METHOD INTERNAL ParseResponsePayload : DINT
VAR_INPUT
  /// Response data
  ResponseData : RobotLibraryResponseDataFB;
  /// Timestamp
  Timestamp    : SystemTime;  
END_VAR
VAR
  /// Parameter count
 _parameterCnt : DINT;
END_VAR
// Table 6-18: Received CMD payload (RC to PLC) of "ReadRobotData"
// --------------------------
// Header
// --------------------------
// Byte 00 : USINT   - ParSeq | State     
// Byte 01 : SINT    - AlarmMessageSeverity    
// Byte 02 : UINT    - AlarmMessageCode HB
// Byte 03 :         - AlarmMessageCode LB
// --------------------------
// Datablock
// --------------------------
// Byte 04 : CHAR  RCManufacturer[0];
// Byte 05 : CHAR  RCManufacturer[1];
// Byte 06 : CHAR  RCManufacturer[2];
// Byte 07 : CHAR  RCManufacturer[3];
// Byte 08 : CHAR  RCManufacturer[4];
// Byte 09 : CHAR  RCManufacturer[5];
// Byte 10 : CHAR  RCManufacturer[6];
// Byte 11 : CHAR  RCManufacturer[7];
// Byte 12 : CHAR  RCManufacturer[8];
// Byte 13 : CHAR  RCManufacturer[9];
// Byte 14 : CHAR  RCManufacturer[10];
// Byte 15 : CHAR  RCManufacturer[11];
// Byte 16 : CHAR  RCManufacturer[12];
// Byte 17 : CHAR  RCManufacturer[13];
// Byte 18 : CHAR  RCManufacturer[14];
// Byte 19 : CHAR  RCManufacturer[15];
// Byte 20 : CHAR  RCManufacturer[16];
// Byte 21 : CHAR  RCManufacturer[17];
// Byte 22 : CHAR  RCManufacturer[18];
// Byte 23 : CHAR  RCManufacturer[19];
// Byte 24 : CHAR  RCOrderID[0];
// Byte 25 : CHAR  RCOrderID[1];
// Byte 26 : CHAR  RCOrderID[2];
// Byte 27 : CHAR  RCOrderID[3];
// Byte 28 : CHAR  RCOrderID[4];
// Byte 29 : CHAR  RCOrderID[5];
// Byte 30 : CHAR  RCOrderID[6];
// Byte 31 : CHAR  RCOrderID[7];
// Byte 32 : CHAR  RCOrderID[8];
// Byte 33 : CHAR  RCOrderID[9];
// Byte 34 : CHAR  RCOrderID[10];
// Byte 35 : CHAR  RCOrderID[11];
// Byte 36 : CHAR  RCOrderID[12];
// Byte 37 : CHAR  RCOrderID[13];
// Byte 38 : CHAR  RCOrderID[14];
// Byte 39 : CHAR  RCOrderID[15];
// Byte 40 : CHAR  RCOrderID[16];
// Byte 41 : CHAR  RCOrderID[17];
// Byte 42 : CHAR  RCOrderID[18];
// Byte 43 : CHAR  RCOrderID[19];
// Byte 44 : CHAR  RCSerialNumber[0];
// Byte 45 : CHAR  RCSerialNumber[1];
// Byte 46 : CHAR  RCSerialNumber[2];
// Byte 47 : CHAR  RCSerialNumber[3];
// Byte 48 : CHAR  RCSerialNumber[4];
// Byte 49 : CHAR  RCSerialNumber[5];
// Byte 50 : CHAR  RCSerialNumber[6];
// Byte 51 : CHAR  RCSerialNumber[7];
// Byte 52 : CHAR  RCSerialNumber[8];
// Byte 53 : CHAR  RCSerialNumber[9];
// Byte 54 : CHAR  RCSerialNumber[10];
// Byte 55 : CHAR  RCSerialNumber[11];
// Byte 56 : CHAR  RCSerialNumber[12];
// Byte 57 : CHAR  RCSerialNumber[13];
// Byte 58 : CHAR  RCSerialNumber[14];
// Byte 59 : CHAR  RCSerialNumber[15];
// Byte 60 : CHAR  RASerialNumber[0];
// Byte 61 : CHAR  RASerialNumber[1];
// Byte 62 : CHAR  RASerialNumber[2];
// Byte 63 : CHAR  RASerialNumber[3];
// Byte 64 : CHAR  RASerialNumber[4];
// Byte 65 : CHAR  RASerialNumber[5];
// Byte 66 : CHAR  RASerialNumber[6];
// Byte 67 : CHAR  RASerialNumber[7];
// Byte 68 : CHAR  RASerialNumber[8];
// Byte 69 : CHAR  RASerialNumber[9];
// Byte 70 : CHAR  RASerialNumber[10];
// Byte 71 : CHAR  RASerialNumber[11];
// Byte 72 : CHAR  RASerialNumber[12];
// Byte 73 : CHAR  RASerialNumber[13];
// Byte 74 : CHAR  RASerialNumber[14];
// Byte 75 : CHAR  RASerialNumber[15];
// Byte 76 : CHAR  RCFirmwareVersion[0];
// Byte 77 : CHAR  RCFirmwareVersion[1];
// Byte 78 : CHAR  RCFirmwareVersion[2];
// Byte 79 : CHAR  RCFirmwareVersion[3];
// Byte 80 : CHAR  RCFirmwareVersion[4];
// Byte 81 : CHAR  RCFirmwareVersion[5];
// Byte 82 : CHAR  RCFirmwareVersion[6];
// Byte 83 : CHAR  RCFirmwareVersion[7];
// Byte 84 : CHAR  RCFirmwareVersion[8];
// Byte 85 : CHAR  RCFirmwareVersion[9];
// Byte 86 : CHAR  RCFirmwareVersion[10];
// Byte 87 : CHAR  RCFirmwareVersion[11];
// Byte 88 : CHAR  RCInterpreterVersion[0];
// Byte 89 : CHAR  RCInterpreterVersion[1];
// Byte 90 : CHAR  RCInterpreterVersion[2];
// Byte 91 : BYTE  Reserved;
// Byte 92 : BYTE  AxisJointUsed;
// Byte 93 : BYTE  AxisExternalUsed;
// Byte 94 : BYTE  AxisJointUnit;
// Byte 95 : BYTE  AxisExternalUnit;
// Byte 96 : BYTE  RCSupportedFunctions[0];
// Byte 97 : BYTE  RCSupportedFunctions[1];
// Byte 98 : BYTE  RCSupportedFunctions[2];
// Byte 99 : BYTE  RCSupportedFunctions[3];
// Byte 100: BYTE  RCSupportedFunctions[4];
// Byte 101: BYTE  RCSupportedFunctions[5];
// Byte 102: BYTE  RCSupportedFunctions[6];
// Byte 103: BYTE  RCSupportedFunctions[7];
// Byte 104: BYTE  RCSupportedFunctions[8];
// Byte 105: BYTE  RCSupportedFunctions[9];
// Byte 106: BYTE  RCSupportedFunctions[10];
// Byte 107: BYTE  RCSupportedFunctions[11];
// Byte 108: BYTE  RCSupportedFunctions[12];
// Byte 109: BYTE  RCSupportedFunctions[13];
// Byte 110: BYTE  RCSupportedFunctions[14];
// Byte 111: BYTE  RCSupportedFunctions[15];
// Byte 112: BYTE  RCSupportedFunctions[16];
// Byte 113: BYTE  RCSupportedFunctions[17];
// Byte 114: BYTE  RCSupportedFunctions[18];
// Byte 115: BYTE  Reserved;
// Byte 116: CHAR  RobotID[0];
// Byte 117: CHAR  RobotID[1];
// Byte 118: CHAR  RobotID[2];
// Byte 119: CHAR  RobotID[3];
// Byte 120: CHAR  RobotID[4];
// Byte 121: CHAR  RobotID[5];
// Byte 122: CHAR  RobotID[6];
// Byte 123: CHAR  RobotID[7];
// Byte 124: CHAR  RobotID[8];
// Byte 125: CHAR  RobotID[9];
// Byte 126: CHAR  RobotID[10];
// Byte 127: CHAR  RobotID[11];
// Byte 128: CHAR  RobotID[12];
// Byte 129: CHAR  RobotID[13];
// Byte 130: CHAR  RobotID[14];
// Byte 131: CHAR  RobotID[15];
// Byte 132: UINT  InterpreterCycleTime HW HB;
// Byte 133:       InterpreterCycleTime HW LB;
// --------------------------

                  
                  // call base implementation to parse the header from payload buffer
ResponseData.PayloadPtr := SUPER^.ParseResponsePayload(ResponseData := ResponseData, Timestamp := Timestamp);

// ST-FIX F100: missing (trailing zero) bytes of the payload are 0, no values of the previous response
SysDepMemSet( pDest := ADR(_response), Value := 0, DataLen := SIZEOF(_response));

// copy parsed header to response
_response.ParSeq               := _rspHeader.ParSeq;
_response.State                := _rspHeader.State;
_response.AlarmMessageSeverity := _rspHeader.AlarmMessageSeverity;
_response.AlarmMessageCode     := _rspHeader.AlarmMessageCode;


// Check payload remaining ? 
IF ( ResponseData.IsPayloadRemaining)
THEN  
  // Get _response.RCManufacturer
  ResponseData.GetDataBlock(pData := ADR(_response.RCManufacturer)      , SIZEOF(_response.RCManufacturer   )   , IsString := TRUE );
  // inc parameter counter
 _parameterCnt := _parameterCnt + 1;
END_IF


// Check payload remaining ? 
IF ( ResponseData.IsPayloadRemaining)
THEN  
  // Get _response.RCOrderID
  ResponseData.GetDataBlock(pData := ADR(_response.RCOrderID)           , SIZEOF(_response.RCOrderID        )   , IsString := TRUE );
  // inc parameter counter
 _parameterCnt := _parameterCnt + 1;
END_IF


// Check payload remaining ? 
IF ( ResponseData.IsPayloadRemaining)
THEN  
  // Get _response.RCSerialNumber
  ResponseData.GetDataBlock(pData := ADR(_response.RCSerialNumber)      , SIZEOF(_response.RCSerialNumber   )   , IsString := TRUE );
  // inc parameter counter
 _parameterCnt := _parameterCnt + 1;
END_IF


// Check payload remaining ? 
IF ( ResponseData.IsPayloadRemaining)
THEN  
  // Get _response.RASerialNumber
  ResponseData.GetDataBlock(pData := ADR(_response.RASerialNumber)      , SIZEOF(_response.RASerialNumber   )   , IsString := TRUE );
  // inc parameter counter
 _parameterCnt := _parameterCnt + 1;
END_IF


// Check payload remaining ? 
IF ( ResponseData.IsPayloadRemaining)
THEN  
  // Get _response.RCFirmwareVersion
  ResponseData.GetDataBlock(pData := ADR(_response.RCFirmwareVersion)   , SIZEOF(_response.RCFirmwareVersion)   , IsString := TRUE );
  // inc parameter counter
 _parameterCnt := _parameterCnt + 1;
END_IF


// Check payload remaining ? 
IF ( ResponseData.IsPayloadRemaining)
THEN  
  // Get _response.RCInterpreterVersion
  // ResponseData.GetDataBlock(pData := ADR(_response.RCInterpreterVersion), SIZEOF(_response.RCInterpreterVersion), IsString := TRUE );

  // This adaption was made because of Stäubli - check with other robot brands...
  
  // Get _response.RCInterpreterVersion
 // ST-FIX F163: the three numbers, the text is made of them
   _response.RCInterpreterVersionNumber.MajorVersion := BYTE_TO_USINT(ResponseData.GetByte());
   _response.RCInterpreterVersionNumber.MinorVersion := BYTE_TO_USINT(ResponseData.GetByte());
   _response.RCInterpreterVersionNumber.PatchVersion := BYTE_TO_USINT(ResponseData.GetByte());
   _response.RCInterpreterVersion := CONCAT(USINT_TO_STRING(_response.RCInterpreterVersionNumber.MajorVersion), '.');
   _response.RCInterpreterVersion := CONCAT(_response.RCInterpreterVersion, USINT_TO_STRING(_response.RCInterpreterVersionNumber.MinorVersion));
   _response.RCInterpreterVersion := CONCAT(_response.RCInterpreterVersion, '.');
   _response.RCInterpreterVersion := CONCAT(_response.RCInterpreterVersion, USINT_TO_STRING(_response.RCInterpreterVersionNumber.PatchVersion));

  // inc parameter counter
 _parameterCnt := _parameterCnt + 1;
END_IF


// Check payload remaining ? 
IF ( ResponseData.IsPayloadRemaining)
THEN  
  // Get _response.Reserve
 _response.Reserve := ResponseData.GetByte(); 
  // inc parameter counter
 _parameterCnt := _parameterCnt + 1;
END_IF


// Check payload remaining ? 
IF ( ResponseData.IsPayloadRemaining)
THEN  
  // Get _response.AxisJointUsed
 _response.AxisJointUsed := ResponseData.GetByte(); 
  // inc parameter counter
 _parameterCnt := _parameterCnt + 1;
END_IF


// Check payload remaining ? 
IF ( ResponseData.IsPayloadRemaining)
THEN  
  // Get _response.AxisExternalUsed
 _response.AxisExternalUsed := ResponseData.GetByte(); 
  // inc parameter counter
 _parameterCnt := _parameterCnt + 1;
END_IF


// Check payload remaining ? 
IF ( ResponseData.IsPayloadRemaining)
THEN  
  // Get _response.AxisJointUnit
 _response.AxisJointUnit := ResponseData.GetByte(); 
  // inc parameter counter
 _parameterCnt := _parameterCnt + 1;
END_IF


// Check payload remaining ? 
IF ( ResponseData.IsPayloadRemaining)
THEN  
  // Get _response.AxisExternalUnit
 _response.AxisExternalUnit := ResponseData.GetByte();
  // inc parameter counter
 _parameterCnt := _parameterCnt + 1;
END_IF


// Check payload remaining ? 
IF ( ResponseData.IsPayloadRemaining)
THEN  
  // Get _response.RCSupportedFunctions
  ResponseData.GetDataBlock(pData := ADR(_response.RCSupportedFunctions), SIZEOF(_response.RCSupportedFunctions), IsString := FALSE );
  // inc parameter counter
 _parameterCnt := _parameterCnt + 1;
END_IF


// Check payload remaining ? 
IF ( ResponseData.IsPayloadRemaining)
THEN  
  // Get _response.Reserve2
 _response.Reserve2 := ResponseData.GetByte(); 
  // inc parameter counter
 _parameterCnt := _parameterCnt + 1;
END_IF


// Check payload remaining ? 
IF ( ResponseData.IsPayloadRemaining)
THEN  
  // Get _response.RobotID
  ResponseData.GetDataBlock(pData := ADR(_response.RobotID)             , SIZEOF(_response.RobotID)             , IsString := TRUE );
  // inc parameter counter
 _parameterCnt := _parameterCnt + 1;
END_IF


// Check payload remaining ? 
IF ( ResponseData.IsPayloadRemaining)
THEN  
  // Get _response.InterpreterCycleTime
 _response.InterpreterCycleTime := ResponseData.GetUint(); // ST-FIX F30 
  // inc parameter counter
 _parameterCnt := _parameterCnt + 1;
END_IF

 
// Create logging
ParseResponsePayloadLog(ResponseData := ResponseData, Timestamp := Timestamp, ParameterCnt := _parameterCnt);
END_METHOD

METHOD INTERNAL ParseResponsePayloadLog
VAR_INPUT
  /// Response data
  ResponseData : RobotLibraryResponseDataFB;
  /// Timestamp
  Timestamp    : SystemTime;  
  /// Parameter count
  ParameterCnt : DINT;
END_VAR
VAR 
  /// internal index for loops
 _idx : DINT;
  /// temporary string
 _tmpStr : STRING;
END_VAR
// Create log entry for Parameter start
CreateLogMessagePara1 ( Timestamp   := Timestamp,
                        MessageType := MessageType.CMD,
                        Severity    := Severity.DEBUG,
                        MessageCode := 0,
                        MessageText := '{1} parameter(s) to parse from the response data:',
                        Para1       := DINT_TO_STRING(ParameterCnt));


// Return if no parameter is remaining...
IF ( ParameterCnt = 0 ) THEN RETURN; END_IF
// dec remaining parameter(s)                        
ParameterCnt := ParameterCnt - 1;
// Create log entry for RCManufacturer
CreateLogMessagePara1 ( Timestamp   := Timestamp,
                        MessageType := MessageType.CMD,
                        Severity    := Severity.DEBUG,
                        MessageCode := 0,
                        MessageText := 'Response.RCManufacturer = {1}',
                        Para1       := _response.RCManufacturer);


// Return if no parameter is remaining...
IF ( ParameterCnt = 0 ) THEN RETURN; END_IF
// dec remaining parameter(s)                        
ParameterCnt := ParameterCnt - 1;
// Create log entry for RCOrderID
CreateLogMessagePara1 ( Timestamp   := Timestamp,
                        MessageType := MessageType.CMD,
                        Severity    := Severity.DEBUG,
                        MessageCode := 0,
                        MessageText := 'Response.RCOrderID = {1}',
                        Para1       := _response.RCOrderID);


// Return if no parameter is remaining...
IF ( ParameterCnt = 0 ) THEN RETURN; END_IF
// dec remaining parameter(s)                        
ParameterCnt := ParameterCnt - 1;
// Create log entry for RCSerialNumber
CreateLogMessagePara1 ( Timestamp   := Timestamp,
                        MessageType := MessageType.CMD,
                        Severity    := Severity.DEBUG,
                        MessageCode := 0,
                        MessageText := 'Response.RCSerialNumber = {1}',
                        Para1       := _response.RCSerialNumber);


// Return if no parameter is remaining...
IF ( ParameterCnt = 0 ) THEN RETURN; END_IF
// dec remaining parameter(s)                        
ParameterCnt := ParameterCnt - 1;
// Create log entry for RASerialNumber
CreateLogMessagePara1 ( Timestamp   := Timestamp,
                        MessageType := MessageType.CMD,
                        Severity    := Severity.DEBUG,
                        MessageCode := 0,
                        MessageText := 'Response.RASerialNumber = {1}',
                        Para1       := _response.RASerialNumber);


// Return if no parameter is remaining...
IF ( ParameterCnt = 0 ) THEN RETURN; END_IF
// dec remaining parameter(s)                        
ParameterCnt := ParameterCnt - 1;
// Create log entry for RCFirmwareVersion
CreateLogMessagePara1 ( Timestamp   := Timestamp,
                        MessageType := MessageType.CMD,
                        Severity    := Severity.DEBUG,
                        MessageCode := 0,
                        MessageText := 'Response.RCFirmwareVersion = {1}',
                        Para1       := _response.RCFirmwareVersion);
                        

// Return if no parameter is remaining...
IF ( ParameterCnt = 0 ) THEN RETURN; END_IF
// dec remaining parameter(s)                        
ParameterCnt := ParameterCnt - 1;
// Create log entry for RCInterpreterVersion
CreateLogMessagePara1 ( Timestamp   := Timestamp,
                        MessageType := MessageType.CMD,
                        Severity    := Severity.DEBUG,
                        MessageCode := 0,
                        MessageText := 'Response.RCInterpreterVersion = {1}',
                        Para1       := _response.RCInterpreterVersion);


// Return if no parameter is remaining...
IF ( ParameterCnt = 0 ) THEN RETURN; END_IF
// dec remaining parameter(s)                        
ParameterCnt := ParameterCnt - 1;
// Create log entry for Reserve
CreateLogMessagePara1 ( Timestamp   := Timestamp,
                        MessageType := MessageType.CMD,
                        Severity    := Severity.DEBUG,
                        MessageCode := 0,
                        MessageText := 'Response.Reserve = {1}',
                        Para1       :=  BYTE_TO_STRING(_response.Reserve));


// Return if no parameter is remaining...
IF ( ParameterCnt = 0 ) THEN RETURN; END_IF
// dec remaining parameter(s)                        
ParameterCnt := ParameterCnt - 1;
// Create log entry for AxisJointUsed
CreateLogMessagePara1 ( Timestamp   := Timestamp,
                        MessageType := MessageType.CMD,
                        Severity    := Severity.DEBUG,
                        MessageCode := 0,
                        MessageText := 'Response.AxisJointUsed = {1}',
                        Para1       :=  BYTE_TO_STRING_BIN(_response.AxisJointUsed));


// Return if no parameter is remaining...
IF ( ParameterCnt = 0 ) THEN RETURN; END_IF
// dec remaining parameter(s)                        
ParameterCnt := ParameterCnt - 1;
// Create log entry for AxisExternalUsed
CreateLogMessagePara1 ( Timestamp   := Timestamp,
                        MessageType := MessageType.CMD,
                        Severity    := Severity.DEBUG,
                        MessageCode := 0,
                        MessageText := 'Response.AxisExternalUsed = {1}',
                        Para1       :=  BYTE_TO_STRING_BIN(_response.AxisExternalUsed));


// Return if no parameter is remaining...
IF ( ParameterCnt = 0 ) THEN RETURN; END_IF
// dec remaining parameter(s)                        
ParameterCnt := ParameterCnt - 1;
// Create log entry for AxisJointUnit
CreateLogMessagePara1 ( Timestamp   := Timestamp,
                        MessageType := MessageType.CMD,
                        Severity    := Severity.DEBUG,
                        MessageCode := 0,
                        MessageText := 'Response.AxisJointUnit = {1}',
                        Para1       :=  BYTE_TO_STRING(_response.AxisJointUnit));


// Return if no parameter is remaining...
IF ( ParameterCnt = 0 ) THEN RETURN; END_IF
// dec remaining parameter(s)                        
ParameterCnt := ParameterCnt - 1;
// Create log entry for AxisExternalUnit
CreateLogMessagePara1 ( Timestamp   := Timestamp,
                        MessageType := MessageType.CMD,
                        Severity    := Severity.DEBUG,
                        MessageCode := 0,
                        MessageText := 'Response.AxisExternalUnit = {1}',
                        Para1       :=  BYTE_TO_STRING(_response.AxisExternalUnit));

FOR _idx := 0 TO 18
do
 _tmpStr := '2#';
 _tmpStr := CONCAT( _tmpStr, BYTE_TO_STRING_BIN(_response.RCSupportedFunctions[_idx]));

  // Return if no parameter is remaining...
  IF ( ParameterCnt = 0 ) THEN RETURN; END_IF
  // dec remaining parameter(s)                        
  ParameterCnt := ParameterCnt - 1;
  // Create log entry for RCSupportedFunctions
  CreateLogMessagePara2 ( Timestamp   := Timestamp,
                          MessageType := MessageType.CMD,
                          Severity    := Severity.DEBUG,
                          MessageCode := 0,
                          MessageText := 'Response.RCSupportedFunctions[{2}] = {1}',
                          Para1       := _tmpStr,
                          Para2       :=  DINT_TO_STRING(_idx));
END_FOR


// Return if no parameter is remaining...
IF ( ParameterCnt = 0 ) THEN RETURN; END_IF
// dec remaining parameter(s)                        
ParameterCnt := ParameterCnt - 1;
// Create log entry for Reserve2
CreateLogMessagePara1 ( Timestamp   := Timestamp,
                        MessageType := MessageType.CMD,
                        Severity    := Severity.DEBUG,
                        MessageCode := 0,
                        MessageText := 'Response.Reserve2 = {1}',
                        Para1       :=  BYTE_TO_STRING(_response.Reserve2));


// Return if no parameter is remaining...
IF ( ParameterCnt = 0 ) THEN RETURN; END_IF
// dec remaining parameter(s)                        
ParameterCnt := ParameterCnt - 1;
// Create log entry for RobotID
CreateLogMessagePara1 ( Timestamp   := Timestamp,
                        MessageType := MessageType.CMD,
                        Severity    := Severity.DEBUG,
                        MessageCode := 0,
                        MessageText := 'Response.RobotID = {1}',
                        Para1       :=  _response.RobotID);


// Return if no parameter is remaining...
IF ( ParameterCnt = 0 ) THEN RETURN; END_IF
// dec remaining parameter(s)                        
ParameterCnt := ParameterCnt - 1;
// Create log entry for InterpreterCycleTime
CreateLogMessagePara1 ( Timestamp   := Timestamp,
                        MessageType := MessageType.CMD,
                        Severity    := Severity.DEBUG,
                        MessageCode := 0,
                        MessageText := 'Response.InterpreterCycleTime = {1}',
                        Para1       :=  UINT_TO_STRING(_response.InterpreterCycleTime));
END_METHOD

METHOD PROTECTED Reset : DINT
VAR_INPUT
END_VAR
Reset := SUPER^.Reset();

Done               := FALSE;
Busy               := FALSE;
CommandBuffered    := FALSE;
END_METHOD

END_FUNCTION_BLOCK

// Library/POUs/_internal/BaseFBs/RobotLibraryBaseExecuteFB
FUNCTION_BLOCK RobotLibraryBaseExecuteFB EXTENDS RobotLibraryBaseFB
// ------------------------------------------------------------------------- 
//  SRCI Robot Library                                                
// ------------------------------------------------------------------------- 
//                                                                           
//  Object:      RobotLibraryBaseFB                                       
//  Author:      Thorsten Brach                                                
//  Date:        2024-08-11
//
//  Description:                                              
//   
//                                                                           
//  Copyright: 
//    (C) 2024 Thorsten Brach. All rights reserved                                                                                                                                            
//             Licensed under the MIT License.
//                                                                           
//  Disclaimer:                                                                           
//    This project is provided without any guarantee and can be used for   
//    private and commercial purposes. Any use is at the user’s 
//    own risk and responsibility.
//
// -------------------------------------------------------------------------
VAR_INPUT
  /// Start of the command at the rising edge
  Execute         : BOOL;
END_VAR
VAR_OUTPUT
  /// The command has been completed successfully
  Done            : BOOL;
  /// FB is being processed
  Busy            : BOOL;
  /// Command is transferred and confirmed by the RC
//  CommandBuffered : BOOL;  
END_VAR


VAR
  /// Rising edge for execute
  {attribute 'hide'}
 _execute_R       : R_TRIG;
  /// Falling edge for execute
  {attribute 'hide'}
 _execute_F       : F_TRIG;
END_VAR
            
          
VAR
  _executeIn : BOOL;
  _executeHold : BOOL;
END_VAR
VAR
  /// ST-FIX F104: rising edge of the Execute input (also while Busy)
  _executeRestart_R : R_TRIG;
END_VAR

// ST-FIX F50: a falling edge of Execute must not cancel the command (spec 5.5.x "Output
// status"): Execute is held internally while Busy; Done/Error/CommandAborted of a command
// whose Execute is already FALSE are shown for one cycle, then the block resets
_executeIn := Execute;
// ST-FIX F104: rising edge of the Execute input also while Busy (Execute is held, F50)
_executeRestart_R(CLK := Execute);
Execute     := Execute OR _executeHold;
SUPER^(AxesGroup := AxesGroup);
_executeHold := Busy;
Execute      := _executeIn;

// Base implementation must be called ! 
METHOD PROTECTED OnCall
VAR_IN_OUT
  /// Robot assignment of function
  AxesGroup         : AxesGroup; 
END_VAR

VAR
  /// internal return value
 _retVal : DINT;
END_VAR
SUPER^.OnCall(AxesGroup := AxesGroup);

// building rising and falling edges
_execute_R( CLK := Execute);
_execute_F( CLK := Execute);


// Check command execution is allowed ?
IF ((     Execute                                ) AND
    ( NOT AxesGroup.State.CMDsEnabled            ) AND
    (     MyType <> 'MC_ExchangeConfigurationFB' ) AND // is part of init sequence
    (     MyType <> 'MC_ReadMessagesFB'          ) AND // is part of init sequence
    (     MyType <> 'MC_ReadRobotDataFB'         ))    // is part of init sequence
THEN
  SetError( ErrorID := RobotLibraryErrorIdEnum.ERR_COMMANDS_NOT_ENABLED, Overwrite := TRUE );
  Error   := TRUE;
  Busy    := FALSE;
END_IF


// On execution started
IF ( _execute_R.Q )
THEN
  OnExecStart(AxesGroup := AxesGroup);
END_IF


// On execution cancel  
IF ( Busy ) AND ( _execute_F.Q ) 
THEN
  // set cancel flag
 _cancel := TRUE;
END_IF

IF ( _cancel )
THEN
  // call Cancel
 _retVal := OnExecCancel(AxesGroup := AxesGroup);
  
  // done or error ?
  IF ( _retVal <> RobotLibraryConstants.RUNNING )
  THEN
    // reset cancel flag
   _cancel := FALSE;
	END_IF
END_IF


// On execution error clear
IF ( Error ) AND ( _execute_F.Q )
THEN
  // set ClearError flag
 _clearError := TRUE;
END_IF

IF ( _clearError )
THEN
 _retVal := OnExecErrorClear(AxesGroup := AxesGroup); 

  // done or error ?
  IF ( _retVal <> RobotLibraryConstants.RUNNING )
  THEN
    // reset ClearError flag
   _clearError := FALSE;
	END_IF
END_IF
END_METHOD

METHOD PROTECTED OnExecCancel : DINT
VAR_IN_OUT
  /// Robot assignment of function
  AxesGroup : AxesGroup; 
END_VAR
VAR
  /// internal return value 
 _retVal    : DINT;
END_VAR
// Create log entry
CreateLogMessagePara1 ( Timestamp   := AxesGroup.State.SystemTime,
                        MessageType := MessageType.CMD,
                        Severity    := Severity.DEBUG,
                        MessageCode := 0,
                        MessageText := 'Execution of {1} cancled ',
                        Para1       := MyType);                 

// try to remove cmd
_retVal := AxesGroup.Acyclic.ActiveCommandRegister.RemoveCmd(_uniqueID);


IF (_retVal = RobotLibraryConstants.OK)
THEN
  // Create log entry
  CreateLogMessagePara1 ( Timestamp   := AxesGroup.State.SystemTime,
                          MessageType := MessageType.CMD,
                          Severity    := Severity.DEBUG,
                          MessageCode := 0,
                          MessageText := '{1} successfully removed from ACR',
                          Para1       := MyType);                 
ELSE
  // Create log entry
  CreateLogMessagePara1 ( Timestamp   := AxesGroup.State.SystemTime,
                          MessageType := MessageType.CMD,
                          Severity    := Severity.DEBUG,
                          MessageCode := 0,
                          MessageText := '{1} was not removed from ACR because execution was already in progress',
                          Para1       := MyType);                 
END_IF


OnExecCancel := Reset();
END_METHOD

METHOD PROTECTED OnExecErrorClear : DINT
VAR_IN_OUT
  /// Robot assignment of function
  AxesGroup : AxesGroup; 
END_VAR
OnExecErrorClear := Reset();
END_METHOD

METHOD PROTECTED OnExecRun : DINT
VAR_IN_OUT
  /// Robot assignment of function
  AxesGroup : AxesGroup; 
END_VAR
END_METHOD

METHOD PROTECTED OnExecStart : DINT
VAR_IN_OUT
  /// Robot assignment of function
  AxesGroup : AxesGroup; 
END_VAR


// ST-FIX F71: Priority (1 = very high ... 4 = low, table 7-1)
IF ( Priority < PriorityLevel.VERY_HIGH )
THEN
  SetError( ErrorID := RobotLibraryErrorIdEnum.ERR_PRIORITY_TOO_HIGH, Overwrite := TRUE );
  // Create log entry
  CreateLogMessage ( Timestamp   := AxesGroup.State.SystemTime,
                     MessageType := MessageType.CMD,
                     Severity    := Severity.ERROR,
                     MessageCode := ErrorID,
                     MessageText := 'Invalid input Priority: higher than VERY_HIGH');
  Error := TRUE;
ELSIF ( Priority > PriorityLevel.LOW )
THEN
  SetError( ErrorID := RobotLibraryErrorIdEnum.ERR_PRIORITY_TOO_LOW, Overwrite := TRUE );
  // Create log entry
  CreateLogMessage ( Timestamp   := AxesGroup.State.SystemTime,
                     MessageType := MessageType.CMD,
                     Severity    := Severity.ERROR,
                     MessageCode := ErrorID,
                     MessageText := 'Invalid input Priority: lower than LOW');
  Error := TRUE;
END_IF
END_METHOD

METHOD PROTECTED OnUpdateStateFlags
VAR_INPUT
  /// Command message state
  State : CmdMessageState;
END_VAR
// Reset State flags
Done := FALSE;

CASE State OF

  // No operation or process is active
  CmdMessageState.EMPTY               :;
  // Created but not yet started
  CmdMessageState.CREATED             :;
  // Buffered and awaiting execution
  CmdMessageState.BUFFERED            :;
  // Buffered in planner for future execution
  CmdMessageState.BUFFERED_IN_PLANNER :;
  // Currently active and in progress
  CmdMessageState.ACTIVE              :;
  // Interrupted and awaiting continuation
  CmdMessageState.INTERRUPTED         :;
  // Requested for abort
  CmdMessageState.ABORT_REQUEST       :;
  // Successfully completed
  CmdMessageState.DONE                : Done := TRUE;
                                        Busy := FALSE;
  // Aborted before completion
  CmdMessageState.ABORTED             : Busy := FALSE;
  // Encountered an error during execution
  CmdMessageState.ERROR               : Error := TRUE;
                                        Busy  := FALSE;
END_CASE
END_METHOD

METHOD PROTECTED Reset : DINT
VAR_INPUT
END_VAR
Reset := SUPER^.Reset();

Done := FALSE;
Busy := FALSE;
END_METHOD

END_FUNCTION_BLOCK

// Library/POUs/_internal/LogFBs/AxesGroupMessageLogFB
FUNCTION_BLOCK AxesGroupMessageLogFB IMPLEMENTS IMessageLogger
// ------------------------------------------------------------------------- 
//  SRCI Robot Library                                                
// ------------------------------------------------------------------------- 
//                                                                           
//  Object:      AxesGroupMessageLogFB                                       
//  Author:      Thorsten Brach                                                
//  Date:        2025-01-05
//
//  Description:                                              
//   
//                                                                           
//  Copyright: 
//    (C) 2025 Thorsten Brach. All rights reserved                                                                                                                                            
//             Licensed under the MIT License.
//                                                                           
//  Disclaimer:                                                                           
//    This project is provided without any guarantee and can be used for   
//    private and commercial purposes. Any use is at the user’s 
//    own risk and responsibility.
//
// -------------------------------------------------------------------------
VAR_INPUT
  /// Logging level
  LogLevel         : LogLevel;
  /// Interface to an external logger
  ExternalLogger   : IMessageLogger;
END_VAR


VAR_OUTPUT
  /// Amount of system log entries
  SystemLogEntries : UINT := 0;
  /// Amount of message log entries
  MessagesEntries  : UINT := 0;
  /// System log
  SystemLogs       : ARRAY[0..RobotLibraryParameter.SYSTEM_LOG_MAX ] OF STRING(RobotLibraryParameter.MESSAGE_TEXT_LEN);
  /// Message Log
  Messages         : ARRAY[0..RobotLibraryParameter.MESSAGE_LOG_MAX] OF AlarmMessage;  
END_VAR

METHOD PUBLIC AddMessageLog
VAR_INPUT
  MessageLog : AlarmMessage;
END_VAR

VAR
  /// internal index
 _idx            : DINT;
  /// internal index to delete
 _idxFound       : DINT;
  /// lowest Severity
 _lowestSeverity : Severity := Severity.FATAL_ERROR;
  /// temporary buffer ( must be one element less than the message log !!! )
 _tmpBuffer      : ARRAY[0..RobotLibraryParameter.MESSAGE_LOG_MAX -1] OF AlarmMessage; 
END_VAR

                  // Check entry must be added ? 
IF (( LogLevel  <= MessageLog.Severity     ) AND
    ( LogLevel  >  LogLevelEnum.DEACTIVATE ))
THEN
  // Check message buffer is full ? 
  IF ( MessagesEntries >= RobotLibraryParameter.MESSAGE_LOG_MAX )
  THEN
    // find lowest Severity
    FOR _idx := 1 TO RobotLibraryParameter.MESSAGE_LOG_MAX
    DO
      // check entry has a lower severity ? 
     _lowestSeverity := MIN( Messages[_idx].Severity, _lowestSeverity );
		END_FOR

    // search for the oldes message with a lower Severity 
    FOR _idx := RobotLibraryParameter.MESSAGE_LOG_MAX TO 1 BY -1
    DO
      // message found ?
      IF (( Messages[_idx].Severity <   MessageLog.Severity ) AND
          ( Messages[_idx].Severity <= _lowestSeverity      ))
      THEN
        // save index to delete 
       _idxFound := _idx;
        EXIT;
			END_IF
		END_FOR
    
    // check message must be deleted ? 
    IF ( _idxFound > 0 )
    THEN
      // shift all messages starting from the found index one position forwards
      FOR _idx := _idxFound TO RobotLibraryParameter.MESSAGE_LOG_MAX -1
      DO
        Messages[_idx] := Messages[_idx +1];
			END_FOR
		END_IF
  END_IF  

  // shift all messages one position backwards
  // shift messages log entries
  SysDepMemCpy( pDest := ADR(_tmpBuffer[0]), pSrc := ADR(  Messages[0]), DataLen := SIZEOF(_tmpBuffer));
  SysDepMemCpy( pDest := ADR(  Messages[1]), pSrc := ADR(_tmpBuffer[0]), DataLen := SIZEOF(_tmpBuffer));
  
  
  // Add new message 
  Messages[0].Timestamp   := MessageLog.Timestamp;           
  Messages[0].MessageType := MessageLog.MessageType;
  Messages[0].Severity    := MessageLog.Severity;
  Messages[0].MessageText := MessageLog.MessageText;
  Messages[0].MessageCode := MessageLog.MessageCode;
  Messages[0].AcrID       := MessageLog.AcrID;   // ST-FIX F74
  Messages[0].CmdType     := MessageLog.CmdType; // ST-FIX F74
  
  // inc message counter
  MessagesEntries := DINT_TO_UINT(LIMIT(0, MessagesEntries + 1, RobotLibraryParameter.MESSAGE_LOG_MAX));
END_IF
END_METHOD

METHOD Public AddMessageLogByParameter
VAR_INPUT
  /// Timestamp
  Timestamp   : SystemTime;
  /// Type of message according to Table 5-48:
  MessageType : MessageType;
  /// Severity of message according to Table 5-49: Debug, Info, Warning, Error, Fatal error
  Severity    : Severity;
  /// Code of messages
  MessageCode : DWORD;
  /// Static text of message
  MessageText : STRING(RobotLibraryParameter.MESSAGE_TEXT_LEN);    
END_VAR

VAR
  /// temporary message 
 _message : AlarmMessage;
END_VAR
_message.Timestamp   := Timestamp;
_message.MessageType := MessageType;
_message.MessageCode := MessageCode;
_message.MessageText := MessageText;
_message.Severity    := Severity;

// Add message to message buffer       
AddMessageLog(_message);
END_METHOD

METHOD PUBLIC AddSystemLog
VAR_INPUT
  /// system log message
  SystemLog : STRING(255);
END_VAR
VAR
  /// internal index
 _idx       : DINT;
  /// internal log message 
 _message   : AlarmMessage;
  /// temporary buffer ( must be one element less than the system log !!! )
 _tmpBuffer : ARRAY[0..RobotLibraryParameter.SYSTEM_LOG_MAX -1] OF STRING(RobotLibraryParameter.MESSAGE_TEXT_LEN);
END_VAR
// shift system log entries
SysDepMemCpy( pDest := ADR(_tmpBuffer[0]), pSrc := ADR(SystemLogs[0]), DataLen := SIZEOF(_tmpBuffer));
SysDepMemCpy( pDest := ADR(SystemLogs[1]), pSrc := ADR(_tmpBuffer[0]), DataLen := SIZEOF(_tmpBuffer));

// Delete CR from system log message
SystemLog := StrReplace(SystemLog, '$R', '');
// Delete LF from system log message          
SystemLog := StrReplace(SystemLog, '$N', '');    
       
// Add System log to buffer 
SystemLogs[0] := SystemLog;
 
// inc SystemLog counter
SystemLogEntries := DINT_TO_UINT(LIMIT(0, SystemLogEntries + 1, RobotLibraryParameter.SYSTEM_LOG_MAX));
END_METHOD

METHOD CheckMessageCodePresent : BOOL
VAR_INPUT
  /// Code of messages
  MessageCode : DWORD;
END_VAR

VAR
  /// internal index for loops
 _idx : DINT;
END_VAR
FOR _idx := 0 TO RobotLibraryParameter.MESSAGE_LOG_MAX
DO
  IF (Messages[_idx].MessageCode = MessageCode)
  THEN
    CheckMessageCodePresent := TRUE;
    RETURN;
	END_IF
END_FOR
END_METHOD

METHOD PUBLIC DeleteMessages
VAR_INPUT
END_VAR
// reset messages
SysDepMemSet(ADR(Messages), 0, SIZEOF(Messages));
// reset message counter
MessagesEntries := 0;
END_METHOD

METHOD DeleteSystemLogs
VAR_INPUT
END_VAR
// reset SystemLogs
SysDepMemSet(ADR(SystemLogs), 0, SIZEOF(SystemLogs));
// reset SystemLogs counter
SystemLogEntries := 0;
END_METHOD

END_FUNCTION_BLOCK

// Library/POUs/_internal/SystemData/AxesGroupSystemDataFB
FUNCTION_BLOCK AxesGroupSystemDataFB 
{attribute 'pack_mode' := '1'} 
// ------------------------------------------------------------------------- 
//  SRCI Robot Library                                                
// ------------------------------------------------------------------------- 
//                                                                           
//  Object:      AxesGroupSystemDataFB                                       
//  Author:      Thorsten Brach                                                
//  Date:        2025-08-31
//
//  Description:                                              
//   
//                                                                           
//  Copyright: 
//    (C) 2025 Thorsten Brach. All rights reserved                                                                                                                                            
//             Licensed under the MIT License.
//                                                                           
//  Disclaimer:                                                                           
//    This project is provided without any guarantee and can be used for   
//    private and commercial purposes. Any use is at the user’s 
//    own risk and responsibility.
//
// -------------------------------------------------------------------------
VAR_INPUT
  /// Pointer to ToolData array
  ToolDataPtr       : POINTER TO Tool;
  /// Lower dimension of ToolData array 
  ToolDataMin       : DINT;
  /// Lower dimension of ToolData array
  ToolDataMax       : DINT;
  /// Amount of ToolData elements in array
  ToolDataCount     : UDINT;

  /// Pointer to LoadData array
  LoadDataPtr       : POINTER TO Load;
  /// Lower dimension of LoadData array 
  LoadDataMin       : DINT;
  /// Lower dimension of LoadData array
  LoadDataMax       : DINT;
  /// Amount of Load elements in array
  LoadDataCount     : UDINT;

  /// Pointer to FrameData array
  FrameDataPtr      : POINTER TO Frame;
  /// Lower dimension of FrameData array 
  FrameDataMin      : DINT;
  /// Lower dimension of FrameData array
  FrameDataMax      : DINT;
  /// Amount of FrameData elements in array
  FrameDataCount    : UDINT;
  
  /// Pointer to WorkAreas array
  WorkAreasPtr      : POINTER TO RobotWorkArea;
  /// Lower dimension of WorkAreas array 
  WorkAreasMin      : DINT;
  /// Lower dimension of WorkAreas array
  WorkAreasMax      : DINT;
  /// Amount of WorkAreas elements in array
  WorkAreasCount    : UDINT;
  
  /// Software limits stored on PLC
  SWLimits          : REFERENCE TO SWLimits;
  /// Default dynamics stored on PLC. For more information refer to 5.5.7
  DefaultDynamics   : REFERENCE TO DefaultDynamics;
  /// Reference dynamics stored on PLC. For more information refer to 5.5.7
  ReferenceDynamics : REFERENCE TO ReferenceDynamics;
END_VAR

METHOD UpdateDefaultDynamics : DINT
VAR_INPUT
  /// Default dynamics values according to Table 6-172.
  DynamicValues : DefaultDynamics;
END_VAR
// Check pointer is vaild ?
IF ( NOT __ISVALIDREF(DefaultDynamics))  
THEN
  RETURN;
END_IF

// Applay new values
DefaultDynamics := DynamicValues;
END_METHOD

METHOD UpdateFrameData : DINT
VAR_INPUT
  /// Reference to BaseFB 
  Caller     : REFERENCE TO RobotLibraryBaseFB;
  /// Current System Time
  SystemTime : SystemTime;
  /// Frame index M
  /// • 0: WCS (default) O
  /// • 1..254: UCS (User frames)
  FrameNo    : USINT;
  /// Frame data (see chapter 5.5.6.2)
  FrameData  : FrameData;
END_VAR


VAR
  /// pointer to frame data
  pFrameData : POINTER TO Frame;  
END_VAR
// Check pointer is vaild ?
IF ( FrameDataPtr = RobotLibraryConstants.NULL_POINTER )
THEN
  RETURN;
END_IF

// Check Frame number is in range ?
IF (( FrameNo < FrameDataMin ) OR
    ( FrameNo > FrameDataMax ))
THEN
  IF ( __ISVALIDREF( Caller ))
  THEN
   // set warning
   Caller.SetWarning( WarningID := RobotLibraryWarningIdEnum.WARN_SAVE_FRAME_FAILED, Overwrite := FALSE);
   
   // Create log entry
   Caller.CreateLogMessagePara1 ( Timestamp   := SystemTime,
                                  MessageType := MessageType.CMD,
                                  Severity    := Severity.WARNING,
                                  MessageCode := Caller.WarningID,
                                  MessageText := 'Save FrameData failed. Index {1} not available in user defined system data',
                                  Para1       :=  USINT_TO_STRING(FrameNo));
  END_IF

  RETURN;
END_IF


// Calculate pointer address for the index of the FrameData Array
pFrameData := FrameDataPtr + (( FrameNo - DINT_TO_UDINT(FrameDataMin)) * SIZEOF(Frame));
// copy frame data to Array index
pFrameData^.Available := TRUE;
pFrameData^.Data := FrameData;
END_METHOD

METHOD UpdateLoadData : DINT
VAR_INPUT
  /// Reference to BaseFB 
  Caller     : REFERENCE TO RobotLibraryBaseFB;
  /// Current System Time
  SystemTime : SystemTime;
  /// Specifies the desired target values that shall be written
  /// Load index
  /// •      0: (default) - Not possible to write
  /// • 1..254: Load data
  LoadNo     : USINT;
  /// Load data (see chapter 5.5.6.4)
  LoadData   : LoadData;
END_VAR


VAR
  /// pointer to load data
  pLoadData : POINTER TO Load;  
END_VAR
// Check pointer is vaild ?
IF ( LoadDataPtr = RobotLibraryConstants.NULL_POINTER )
THEN
  RETURN;
END_IF

// Check Load number is in range ?
IF (( LoadNo < LoadDataMin ) OR
    ( LoadNo > LoadDataMax ))
THEN
  IF ( __ISVALIDREF( Caller ))
  THEN
   // set warning
   Caller.SetWarning( WarningID := RobotLibraryWarningIdEnum.WARN_SAVE_LOAD_FAILED, Overwrite := FALSE);
   
   // Create log entry
   Caller.CreateLogMessagePara1 ( Timestamp   := SystemTime,
                                  MessageType := MessageType.CMD,
                                  Severity    := Severity.WARNING,
                                  MessageCode := Caller.WarningID,
                                  MessageText := 'Save LoadData failed. Index {1} not available in user defined system data',
                                  Para1       :=  USINT_TO_STRING(LoadNo));
  END_IF

  RETURN;
END_IF


// Calculate pointer address for the index of the LoadData Array
pLoadData := LoadDataPtr + (( LoadNo - DINT_TO_UDINT(LoadDataMin)) * SIZEOF(Load));
// copy load data to Array index
pLoadData^.Available := TRUE;
pLoadData^.Data := LoadData;
END_METHOD

METHOD UpdateReferenceDynamics : DINT
VAR_INPUT
  /// Reference dynamics values according to Table 6-158.
  DynamicValues : ReferenceDynamics;
END_VAR
// Check pointer is vaild ?
IF ( NOT __ISVALIDREF(ReferenceDynamics))  
THEN
  RETURN;
END_IF

// Applay new values
ReferenceDynamics := DynamicValues;
END_METHOD

METHOD UpdateSWLimits : DINT
VAR_INPUT
  /// Limits for joints and external axes according to Table 6-197.
  LimitValues : SWLimits;
END_VAR
// Check pointer is vaild ?
IF ( NOT __ISVALIDREF(SWLimits))  
THEN
  RETURN;
END_IF

// Applay new values
SWLimits := LimitValues;
END_METHOD

METHOD UpdateToolData : DINT
VAR_INPUT
  /// Reference to BaseFB 
  Caller     : REFERENCE TO RobotLibraryBaseFB;
  /// Current System Time
  SystemTime : SystemTime;
  /// Tool index
  /// •      0: Flange (default) Not possible to change
  /// • 1..254: Tool Frame
  ToolNo     : USINT;
  /// Tool data (see chapter 5.5.6.3)
  ToolData   : ToolData;
END_VAR


VAR
  /// pointer to tool data
  pToolData : POINTER TO Tool;  
END_VAR
// Check pointer is vaild ?
IF ( ToolDataPtr = RobotLibraryConstants.NULL_POINTER )
THEN
  RETURN;
END_IF

// Check Tool number is in range ?
IF (( ToolNo < ToolDataMin ) OR
    ( ToolNo > ToolDataMax ))
THEN
  IF ( __ISVALIDREF( Caller ))
  THEN
   // set warning
   Caller.SetWarning( WarningID := RobotLibraryWarningIdEnum.WARN_SAVE_TOOL_FAILED, Overwrite := FALSE);
   
   // Create log entry
   Caller.CreateLogMessagePara1 ( Timestamp   := SystemTime,
                                  MessageType := MessageType.CMD,
                                  Severity    := Severity.WARNING,
                                  MessageCode := Caller.WarningID,
                                  MessageText := 'Save ToolData failed. Index {1} not available in user defined system data',
                                  Para1       :=  USINT_TO_STRING(ToolNo));
  END_IF

  RETURN;
END_IF

// ST-FIX F81: copy the tool into the ToolData array (was commented out)
// Calculate pointer address for the index of the ToolData Array
pToolData := ToolDataPtr + (( ToolNo - DINT_TO_UDINT(ToolDataMin)) * SIZEOF(Tool));
// copy tool data to Array index
pToolData^.Available := TRUE;
pToolData^.Data := ToolData;
END_METHOD

METHOD UpdateWorAreas : DINT
VAR_INPUT
  /// Reference to BaseFB 
  Caller       : REFERENCE TO RobotLibraryBaseFB;
  /// Current System Time
  SystemTime   : SystemTime;
  /// Index of the robot work area
  /// • 0 (default)..254
  WorkAreaNo   : USINT;
  /// Data specific to the work area requested by Index.
  WorkAreaData : RobotWorkAreaData;
END_VAR
VAR
  /// pointer to WorkArea
  pWorkAreaData : POINTER TO RobotWorkArea;  
END_VAR
// Check pointer is vaild ?
IF ( WorkAreasPtr = RobotLibraryConstants.NULL_POINTER )
THEN
  RETURN;
END_IF

// Check WorkArea number is in range ?
IF (( WorkAreaNo < WorkAreasMin ) OR
    ( WorkAreaNo > WorkAreasMax ))
THEN
  IF ( __ISVALIDREF( Caller ))
  THEN
   // set warning
   Caller.SetWarning( WarningID := RobotLibraryWarningIdEnum.WARN_SAVE_WORKAREA_FAILED, Overwrite := FALSE);
   
   // Create log entry
   Caller.CreateLogMessagePara1 ( Timestamp   := SystemTime,
                                  MessageType := MessageType.CMD,
                                  Severity    := Severity.WARNING,
                                  MessageCode := Caller.WarningID,
                                  MessageText := 'Save WorkArea failed. Index {1} not available in user defined system data',
                                  Para1       :=  USINT_TO_STRING(WorkAreaNo));
  END_IF

  RETURN;
END_IF


// Calculate pointer address for the index of the WorkArea Array
pWorkAreaData := WorkAreasPtr + (( WorkAreaNo - DINT_TO_UDINT(WorkAreasMin)) * SIZEOF(RobotWorkArea));
// copy WorkArea to Array index
pWorkAreaData^.Available := TRUE;
pWorkAreaData^.Data := WorkAreaData;
END_METHOD

END_FUNCTION_BLOCK

// Library/POUs/_internal/ActiveCommandRegisterFB
FUNCTION_BLOCK ActiveCommandRegisterFB EXTENDS RobotLibraryLogFB
// ------------------------------------------------------------------------- 
//  SRCI Robot Library                                                
// ------------------------------------------------------------------------- 
//                                                                           
//  Object:      ActiveCommandRegisterFB                                       
//  Author:      Thorsten Brach                                                
//  Date:        2024-06-01
//
//  Description:                                              
//   
//                                                                           
//  Copyright: 
//    (C) 2024 Thorsten Brach. All rights reserved                                                                                                                                            
//             Licensed under the MIT License.
//                                                                           
//  Disclaimer:                                                                           
//    This project is provided without any guarantee and can be used for   
//    private and commercial purposes. Any use is at the user’s 
//    own risk and responsibility.
//
// -------------------------------------------------------------------------
VAR_INPUT
  /// Active Command Register
  Register            : ARRAY [1..RobotLibraryParameter.ACTIVE_CMD_REGISTER_ENTRIES_MAX] OF AxesGroupAcyclicAcrEntry;
  /// System Time
  SystemTime          : SystemTime;
  /// usable size of the arc register
  RegisterSize        : DINT := RobotLibraryParameter.ACTIVE_CMD_REGISTER_ENTRIES_MAX;
END_VAR

VAR_OUTPUT
  /// Execution Order List 
  ExecutionOrderList    : ARRAY [1..RobotLibraryParameter.ACTIVE_CMD_REGISTER_ENTRIES_MAX] OF DINT;
  /// Current amount of used registers
  CurrentAcrUsageCount  : DINT;  
  /// Current percent of used registers
  CurrentAcrUsagePercent : REAL;    
END_VAR


VAR
  /// temporarty Active Command Register
  TmpRegister                 : ARRAY [1..RobotLibraryParameter.ACTIVE_CMD_REGISTER_ENTRIES_MAX] OF AxesGroupAcyclicAcrEntry;
  /// last used unique ID 
  LastUniqueID                : UINT;
  /// Warning for ACR usage at 80%
  WarningAcrUsage             : R_TRIG;
END_VAR

VAR CONSTANT
  /// Active command
  ACTIVE_CMD           : UDINT := 1;
  /// Buffered command
  BUFFER_CMD           : UDINT := 2;
  /// Empty ACR entry
  EMPTY_ACR_ENTRY      : AxesGroupAcyclicAcrEntry := (State := ActiveCommandRegisterState.IS_FREE);
  /// Empty command entry
  EMPTY_CMD_ENTRY      : AxesGroupAcyclicAcrEntryCmdBuffer := (State := BufferStateCmd.EMPTY);  
  /// constant for byte index of priority in payload 
  PRIORITY_IDX         : BYTE := 3;  
  /// bitmask to mask the priority out of the halfbyte
  PRIORITY_BIT_MASK    : BYTE := 2#000_1111;   
END_VAR

ManageRegister();

UpdateExecutionOrderList();

METHOD PUBLIC AddCmd : UDINT
VAR_INPUT
  /// Pointer to the corresponding command-FB to enable a callback mechanism
  pCommandFB        : POINTER TO RobotLibraryBaseFB;
END_VAR

VAR
  /// internal index for loops
 _regIdx            : DINT;
  /// internal command type 
 _cmdType           : CmdType;
  /// log message
 _messageLog        : AlarmMessage;  
  /// flag for free register found
 _freeRegisterFound : BOOL;
  /// internal Acr error 
 _errorAcrEntry     : WORD := RobotLibraryErrorIdEnum.ERR_NO_FREE_ACR_ENTRY;  
END_VAR

                  // ST-FIX F48: a command with a parameter error of the block is not added
IF ( pCommandFB <> 0 )
THEN
  IF (( pCommandFB^.ErrorID = RobotLibraryErrorIdEnum.ERR_INVALID_PARAM_EXECUTION_MODE ) OR
      ( pCommandFB^.ErrorID = RobotLibraryErrorIdEnum.ERR_PROCESSINGMODE_NOT_DEFINED   ))
  THEN
    AddCmd := 0;
    RETURN;
  END_IF
END_IF

// calculate the used length of the ACR 
FOR _regIdx := 1 TO RegisterSize
DO
  IF ( Register[_regIdx].State = ActiveCommandRegisterState.IS_FREE )
  THEN
    Register[_regIdx].State      := ActiveCommandRegisterState.IS_PROCESSING;
    Register[_regIdx].UniqueID   := DINT_TO_UINT(_regIdx);
    Register[_regIdx].pCommandFB := pCommandFB;

    // check pointer to command FB
    IF ( Register[_regIdx].pCommandFB <> RobotLibraryConstants.NULL_POINTER )
    THEN
      Register[_regIdx].Command[RobotLibraryConstants.ACTIVE_CMD].Timestamp  := SystemTime;

      Register[_regIdx].Command[RobotLibraryConstants.ACTIVE_CMD].Payload    := pCommandFB^.CommandData.Payload; 
      Register[_regIdx].Command[RobotLibraryConstants.ACTIVE_CMD].PayloadLen := pCommandFB^.CommandData.PayloadLen;
      Register[_regIdx].Command[RobotLibraryConstants.ACTIVE_CMD].PayLoadPtr := 0;
      Register[_regIdx].Command[RobotLibraryConstants.ACTIVE_CMD].State      := BufferStateCmd.CREATED;
    END_IF
  
    // set flag for free register found
   _freeRegisterFound := TRUE;
    
    // Increment Current used register counter
    CurrentAcrUsageCount := CurrentAcrUsageCount + 1;
    
    // return Unique ID
    AddCmd := Register[_regIdx].UniqueID;

    // Get CmdType from payload
    SysDepMemCpy( pDest := ADR(_cmdType), pSrc := ADR(pCommandFB^.CommandData.Payload), DataLen := SIZEOF(_cmdType));
    
    // Create log entry
    CreateLogMessagePara2 ( Timestamp   := SystemTime,
                            MessageType := MessageType.CMD,
                            Severity    := Severity.INFO,
                            MessageCode := 0,
                            MessageText := 'ACR-ID [{1}]: Added  Command-Payload of CmdType <{2}>',
                            Para1       :=  DINT_TO_STRING(_regIdx),
                            Para2       :=  CMD_TYPE_TO_STRING(SwapUint(_cmdType)));
    EXIT;
  END_IF
END_FOR

// Check a free register could be found ? 
IF ( NOT _freeRegisterFound )
THEN
  // set error in Command FB   
  IF ( pCommandFB <> RobotLibraryConstants.NULL_POINTER )
  THEN
    SysDepMemCpy( pDest   := ADR   ( pCommandFB^.ErrorID ), 
                  pSrc    := ADR   ( _errorAcrEntry      ),
                  DataLen := SIZEOF( _errorAcrEntry      )); 
  END_IF


  // Create log entry
  CreateLogMessagePara1 ( Timestamp   := SystemTime,
                          MessageType := MessageType.CMD,
                          Severity    := Severity.FATAL_ERROR,
                          MessageCode := 0,
                          MessageText := 'Not possible to add CMD <{1}> to ACR - NO FREE REGISTER FOUND ! -> STOPPING SRCI INTERFACE...',
                          Para1       :=  CMD_TYPE_TO_STRING(SwapUint(_cmdType)));                          
END_IF
END_METHOD

METHOD AddRsp : UDINT
VAR_INPUT
  /// Response
  Rsp : TelegramRobToPlcFragment;
END_VAR
VAR
  /// internal index for loops
 _Idx             : DINT;
  /// internal registen index
 _regIdx          : DINT;
  /// internal command type
 _cmdType         : CmdType;
  /// internal FragmentAction
 _fragmentAction  :  FragmentAction;
  /// internal command message state
 _cmdMessageState : CmdMessageState;
  /// internal flag for CmdID found
 _found           : BOOL;
END_VAR

                  FOR _regIdx := 1 TO RegisterSize
DO
  IF ( Register[_regIdx].UniqueID = Rsp.Header.CmdID )
  THEN
    // CmdID was found in the ACR
   _found := TRUE;
    // convert to fragment action 
   _fragmentAction := ByteToFragmentAction(Rsp.Header.FragmentAction);

    // delete response 
    IF ( _fragmentAction.Clear )
    THEN
      SysDepMemSet( pDest := ADR(Register[_regIdx].Response[ACTIVE_CMD]), Value := 0, DataLen := SIZEOF(Register[_regIdx].Response[ACTIVE_CMD]));
    END_IF
                       
    // add payload to response
    FOR _idx := Rsp.Header.PayloadPointer TO  Rsp.Header.PayloadPointer + Rsp.Header.PayloadLength -1
    DO
      Register[_regIdx].Response[ACTIVE_CMD].Timestamp     := SystemTime;
      Register[_regIdx].Response[ACTIVE_CMD].State         := BufferStateRsp.RECEIVING;
      Register[_regIdx].Response[ACTIVE_CMD].PayloadLen    := Register[_regIdx].Response[ACTIVE_CMD].PayloadLen + 1;
      Register[_regIdx].Response[ACTIVE_CMD].Payload[_idx] := Rsp.Command.Payload[_idx];
    END_FOR

    // Get current message state 
   _cmdMessageState := GetHalfeByteLo    (Value  := Register[_regIdx].Response[ACTIVE_CMD].Payload[0]);
    // Get command type from payload
   _cmdType         := CombineBytesToUint(HiByte := Register[_regIdx].Command [ACTIVE_CMD].Payload[0],
                                          LoByte := Register[_regIdx].Command [ACTIVE_CMD].Payload[1]);

    // Create log entry
    CreateLogMessagePara3 ( Timestamp   := SystemTime,
                            MessageType := MessageType.CMD,
                            Severity    := Severity.INFO,
                            MessageCode := 0,
                            MessageText := 'ACR-ID [{1}]: Added Response-Payload of CmdType <{2}> with State = {3}',
                            Para1       :=  DINT_TO_STRING(_regIdx),
                            Para2       :=  CMD_TYPE_TO_STRING(_cmdType),
                            Para3       :=  CMD_MESSAGE_STATE_TO_STRING(_cmdMessageState));

    IF ( _fragmentAction.Complete )
    THEN
      // set response state
      Register[_regIdx].Response[ACTIVE_CMD].State := BufferStateRsp.RECEIVED;      
     
      // Check current message state and tag the register state as IS_FINAL, if needed 
      IF ( _cmdMessageState >= CmdMessageState.DONE) 
      THEN
        Register[_regIdx].State := ActiveCommandRegisterState.IS_FINAL;
        
        // get command type from payload
       _cmdType := CombineBytesToUint(HiByte := Register[_regIdx].Command[ACTIVE_CMD].Payload[0],
                                      LoByte := Register[_regIdx].Command[ACTIVE_CMD].Payload[1]);

        // Create log entry
        CreateLogMessagePara3( Timestamp   := SystemTime,
                               MessageType := MessageType.CMD,
                               Severity    := Severity.INFO,
                               MessageCode := 0,
                               MessageText := 'ACR-ID [{1}]: Detected Response-Payload of CmdType <{2}> has reached final state <{3}>',
                               Para1       :=  DINT_TO_STRING(_regIdx),
                               Para2       :=  CMD_TYPE_TO_STRING(_cmdType),
                               Para3       :=  CMD_MESSAGE_STATE_TO_STRING(_cmdMessageState));
                               
        // Exit the loop
      END_IF      
    END_IF
    
    
    // Check Response received complete ? 
    IF ( Register[_regIdx].Response[ACTIVE_CMD].State = BufferStateRsp.RECEIVED)
    THEN
      // update state
      Register[_regIdx].Response[ACTIVE_CMD].State := BufferStateRsp.PROCESSED;
      // callback CommandFB    
      Register[_regIdx].pCommandFB^.CallBack(RspData := Register[_regIdx].Response[ACTIVE_CMD],TimeStamp := SystemTime);    
    END_IF
    
    EXIT;
  END_IF
END_FOR


// Check CmdID was found in the ACR ? 
IF ( NOT _found )
THEN
  // Create log entry
  CreateLogMessagePara2 ( Timestamp   := SystemTime,
                          MessageType := MessageType.CMD,
                          Severity    := Severity.WARNING,
                          MessageCode := 0,
                          MessageText := 'ACR-ID [?]: Response-Payload of CmdID <{1}> with State = {2} received, but no matching ACR entry found',
                          Para1       :=  UINT_TO_STRING(Rsp.Header.CmdID),
                          Para2       :=  CMD_MESSAGE_STATE_TO_STRING(_cmdMessageState));
END_IF
END_METHOD

METHOD FB_init : BOOL
VAR_INPUT
  bInitRetains : BOOL; // if TRUE, the retain variables are initialized (warm start / cold start)
  bInCopyCode : BOOL;  // if TRUE, the instance afterwards gets moved into the copy code (online change)
END_VAR
MyType := 'ActiveCommandRegisterFB';
END_METHOD

METHOD PRIVATE ManageRegister
VAR
  /// internal index
 _regIdx          : DINT;
  /// internal command type
 _cmdType         : CmdType;
  /// internal command message state
 _cmdMessageState : CmdMessageState; 
END_VAR
FOR _regIdx := 1 TO RegisterSize
DO
  // Check pointer to command FB is valid ? 
  IF ( Register[_regIdx].pCommandFB <> RobotLibraryConstants.NULL_POINTER) 
  THEN
  
    // Check apply Cmd parameter update ?  
    IF (( Register[_regIdx].Command[ACTIVE_CMD].State = BufferStateCmd.PROCESSED        ) AND
        ( Register[_regIdx].Command[BUFFER_CMD].State = BufferStateCmd.UPDATE_AVAILABLE ))
    THEN
      Register[_regIdx].Command[ACTIVE_CMD] := Register[_regIdx].Command[BUFFER_CMD];
      Register[_regIdx].Command[BUFFER_CMD] := EMPTY_CMD_ENTRY;
  
      // get command type from payload
     _cmdType := CombineBytesToUint(HiByte := Register[_regIdx].Command[ACTIVE_CMD].Payload[0],
                                    LoByte := Register[_regIdx].Command[ACTIVE_CMD].Payload[1]);
  
      // Create log entry
      CreateLogMessagePara2 ( Timestamp   := SystemTime,
                              MessageType := MessageType.CMD,
                              Severity    := Severity.INFO,
                              MessageCode := 0,
                              MessageText := 'ACR-ID [{1}]: Moved BUFFER_CMD to ACTIVE_CMD, CmdType <{2}>',
                              Para1       :=  DINT_TO_STRING(_regIdx),
                              Para2       :=  CMD_TYPE_TO_STRING(_cmdType));
  
    END_IF
    
    (*
    // Check Response received ? 
    IF ( Register[_regIdx].Response[ACTIVE_CMD].State = BufferStateRsp.RECEIVED)
    THEN
      // update state
      Register[_regIdx].Response[ACTIVE_CMD].State := BufferStateRsp.PROCESSED;
      // callback CommandFB    
      Register[_regIdx].pCommandFB^.CallBack(RspData := Register[_regIdx].Response[ACTIVE_CMD],TimeStamp := SystemTime);    
    END_IF
    *)
    
    // delete entries with State.IS_Final 
    IF ( Register[_regIdx].State = ActiveCommandRegisterState.IS_FINAL )
    THEN
      // get command type from payload
     _cmdType := CombineBytesToUint(HiByte := Register[_regIdx].Command[ACTIVE_CMD].Payload[0],
                                    LoByte := Register[_regIdx].Command[ACTIVE_CMD].Payload[1]);
  
      // Get current message state 
     _cmdMessageState := GetHalfeByteLo(Value := Register[_regIdx].Response[ACTIVE_CMD].Payload[0]);

  
      // Create log entry
      CreateLogMessagePara3( Timestamp   := SystemTime,
                             MessageType := MessageType.CMD,
                             Severity    := Severity.INFO,
                             MessageCode := 0,
                             MessageText := 'ACR-ID [{1}]: Deleted ACR-Entry of CmdType <{2}> with State = {3}, because of Final-State was reached',
                             Para1       :=  DINT_TO_STRING(_regIdx),
                             Para2       :=  CMD_TYPE_TO_STRING(_cmdType),
                             Para3       :=  CMD_MESSAGE_STATE_TO_STRING(_cmdMessageState));
  
                             
      // delete register entry                              
      Register[_regIdx] := EMPTY_ACR_ENTRY;

      // decrement current used register counter
      CurrentAcrUsageCount := CurrentAcrUsageCount - 1;                           
    END_IF
  END_IF
END_FOR


// Calculate percent of register usage
IF ( CurrentAcrUsageCount > 0)
THEN
  CurrentAcrUsagePercent :=  (DINT_TO_REAL(CurrentAcrUsageCount) / DINT_TO_REAL(RegisterSize)) * 100.0;
ELSE
  CurrentAcrUsagePercent := 0.0;
END_IF

// build rising edge for arc usage over 80% 
WarningAcrUsage( CLK := CurrentAcrUsagePercent > RobotLibraryParameter.ACR_USAGE_WARNING_LIMIT );

IF ( WarningAcrUsage.Q )
THEN
  // Create log entry
  CreateLogMessagePara4( Timestamp   := SystemTime,
                         MessageType := MessageType.CMD,
                         Severity    := Severity.WARNING,
                         MessageCode := 0,
                         MessageText := 'ACR Register usage has reached the warning limit ({1}): {2}/{3} = {4}%',
                         Para1       :=  REAL_TO_STRING(RobotLibraryParameter.ACR_USAGE_WARNING_LIMIT),
                         Para2       :=  DINT_TO_STRING(CurrentAcrUsageCount),
                         Para3       :=  DINT_TO_STRING(RegisterSize),
                         Para4       :=  REAL_TO_STRING(CurrentAcrUsagePercent));  
END_IF
END_METHOD

PROPERTY PUBLIC NotifyParameterChanged : UDINT
SET
VAR
  /// internal register index
 _regIdx  : DINT;
  /// internal command type
 _cmdType : CmdType;
END_VAR
FOR _regIdx := 1 TO RobotLibraryParameter.ACTIVE_CMD_REGISTER_ENTRIES_MAX
DO
  // check unique ID found ?
  IF ( Register[_regIdx].UniqueID = NotifyParameterChanged )
  THEN  
    // ST-FIX F114: a parameter change before the command is sent (state CREATED) must not turn the new
    // command into a parameter update (it was never sent): the command keeps the parameters of the rising edge
    IF ( Register[_regIdx].Command[ACTIVE_CMD].State = BufferStateCmd.CREATED )
    THEN
      // Create log entry
      CreateLogMessagePara1 ( Timestamp   := SystemTime,
                              MessageType := MessageType.CMD,
                              Severity    := Severity.INFO,
                              MessageCode := 0,
                              MessageText := 'ACR-ID [{1}]: Cmd-Parameter changed before the command was sent -> ignored',
                              Para1       :=  DINT_TO_STRING(_regIdx));
    ELSIF (( Register[_regIdx].Command[ACTIVE_CMD].State <> BufferStateCmd.SENDING   ) AND
           ( Register[_regIdx].Command[ACTIVE_CMD].State <> BufferStateCmd.PROCESSED ))
    THEN
      // Check pointer is valid ? 
      IF ( Register[_regIdx].pCommandFB <> RobotLibraryConstants.NULL_POINTER )
      THEN
        // add to send register
        Register[_regIdx].Command[ACTIVE_CMD].Timestamp  := SystemTime;
        Register[_regIdx].Command[ACTIVE_CMD].State      := BufferStateCmd.UPDATE_AVAILABLE;
        Register[_regIdx].Command[ACTIVE_CMD].Payload    := Register[_regIdx].pCommandFB^.CommandData.Payload;
        Register[_regIdx].Command[ACTIVE_CMD].PayloadLen := Register[_regIdx].pCommandFB^.CommandData.PayloadLen;

        // get command type from payload
       _cmdType := CombineBytesToUint(HiByte := Register[_regIdx].pCommandFB^.CommandData.Payload[0],
                                      LoByte := Register[_regIdx].pCommandFB^.CommandData.Payload[1]);
        
        // Create log entry
        CreateLogMessagePara2 ( Timestamp   := SystemTime,
                                MessageType := MessageType.CMD,
                                Severity    := Severity.INFO,
                                MessageCode := 0,
                                MessageText := 'ACR-ID [{1}]: Updated Cmd-Parameter of CmdType <{2}> -> written to ACTIVE_CMD Index',
                                Para1       :=  DINT_TO_STRING(_regIdx),
                                Para2       :=  CMD_TYPE_TO_STRING(_cmdType));
      END_IF
    ELSE
      // Check pointer is valid ? 
      IF ( Register[_regIdx].pCommandFB <> RobotLibraryConstants.NULL_POINTER )
      THEN
        // add to buffer register
        Register[_regIdx].Command[BUFFER_CMD].Timestamp  := SystemTime;
        Register[_regIdx].Command[BUFFER_CMD].State      := BufferStateCmd.UPDATE_AVAILABLE;
        Register[_regIdx].Command[BUFFER_CMD].Payload    := Register[_regIdx].pCommandFB^.CommandData.Payload;
        Register[_regIdx].Command[BUFFER_CMD].PayloadLen := Register[_regIdx].pCommandFB^.CommandData.PayloadLen;

        // get command type from payload
       _cmdType := CombineBytesToUint(HiByte := Register[_regIdx].pCommandFB^.CommandData.Payload[0],
                                      LoByte := Register[_regIdx].pCommandFB^.CommandData.Payload[1]);
        
        // Create log entry
        CreateLogMessagePara2 ( Timestamp   := SystemTime,
                                MessageType := MessageType.CMD,
                                Severity    := Severity.INFO,
                                MessageCode := 0,
                                MessageText := 'ACR-ID [{1}]: Updated Cmd-Parameter of CmdType <{2}> -> written to BUFFER_CMD Index',
                                Para1       :=  DINT_TO_STRING(_regIdx),
                                Para2       :=  CMD_TYPE_TO_STRING(_cmdType));
      END_IF
    END_IF
    
    
  END_IF
END_FOR
END_SET
END_PROPERTY

METHOD PUBLIC OnOnlineChange : DINT
VAR_INPUT
  /// unique ID 
  UniqueID     : UDINT;
  /// Pointer to the corresponding command-FB to enable a callback mechanism
  pCommandFB   : POINTER TO RobotLibraryBaseFB;
END_VAR

VAR
  /// internal index for loops
 _regIdx : DINT;
END_VAR
OnOnlineChange := -1;

// Check command FB pointer is valid ?
IF ( pCommandFB <> RobotLibraryConstants.NULL_POINTER)
THEN
  FOR _regIdx := 1 TO RegisterSize
  DO
    // check unique ID found ?
    IF ( Register[_regIdx].UniqueID = UniqueID ) 
    THEN  
      // update pointer to command FB
      Register[_regIdx].pCommandFB := pCommandFB;
      // Return result OK
      OnOnlineChange := RobotLibraryConstants.OK;
      EXIT;
    END_IF
  END_FOR
END_IF
END_METHOD

METHOD PUBLIC RemoveCmd : DINT
VAR_INPUT
 /// unique ID
 UniqueID : UDINT;  
END_VAR

VAR
  /// internal index
 _regIdx : DINT;
  /// internal command type 
 _cmdType : CmdType;
END_VAR
RemoveCmd := RobotLibraryConstants.HAS_ERROR;


IF (UniqueID = 0)
THEN
  UniqueID := UniqueID;
END_IF

FOR _regIdx := 1 TO RegisterSize
DO
  // check unique ID found and not yet sended ?
  IF (( Register[_regIdx].UniqueID                  = UniqueID                        ) AND
      ( Register[_regIdx].Command[ACTIVE_CMD].State < BufferStateCmd.UPDATE_AVAILABLE ))       
  THEN
    // Get CmdType from payload
    SysDepMemCpy( pDest := ADR(_cmdType), pSrc := ADR(Register[_regIdx].Command[ACTIVE_CMD].Payload), DataLen := SIZEOF(_cmdType));
    // delete register entry
    SysDepMemSet(pDest := ADR(Register[_regIdx]), Value := 0 , DataLen := SIZEOF(Register[_regIdx]));
    // decrement current used register counter
    CurrentAcrUsageCount := CurrentAcrUsageCount - 1;
    // Command successfull removed
    RemoveCmd := RobotLibraryConstants.OK;    
    
    
    // Create log entry
    CreateLogMessagePara2 (  Timestamp   := SystemTime,
                             MessageType := MessageType.CMD,
                             Severity    := Severity.INFO,
                             MessageCode := 0,
                             MessageText := 'ACR-ID [{1}]: Removed CmdType <{2}>',
                             Para1       :=  DINT_TO_STRING(_regIdx),                 
                             Para2       :=  CMD_TYPE_TO_STRING(SwapUint(_cmdType)));
    EXIT;
  END_IF
END_FOR
END_METHOD

METHOD PUBLIC Reset
SysDepMemSet( ADR(Register), 0, SIZEOF(Register));              

CurrentAcrUsageCount   := 0;
CurrentAcrUsagePercent := 0.0;


// Create log entry
CreateLogMessagePara1 ( Timestamp   := SystemTime,
                        MessageType := MessageType.CMD,
                        Severity    := Severity.INFO,
                        MessageCode := 0,
                        MessageText := 'ACR Registers has been reset and all entries deleted by Reset method call',
                        Para1       :=  '');
END_METHOD

METHOD PRIVATE UpdateExecutionOrderList
VAR
  /// temporary Active Command Register entry
  TmpRegisterEntry : AxesGroupAcyclicAcrEntry;
  /// temporary index
  TmpIndex         : DINT;
  /// internal index
  i                : DINT;  
  /// internal index
  j                : DINT;  
END_VAR
// Reset temporary register
SysDepMemSet(pDest := ADR(TmpRegister)       , Value := 0, DataLen := SIZEOF(TmpRegister));
// Reset Execution Order List
SysDepMemSet(pDest := ADR(ExecutionOrderList), Value := 0, DataLen := SIZEOF(ExecutionOrderList));
// pre-set temporary register index 
j := 1;

FOR i := 1 TO RegisterSize
DO
  // add only entries which are not in status free and where datas must be processed
  IF (( Register[i].State                      > ActiveCommandRegisterState.IS_FREE ) AND
      ( Register[i].Command[ACTIVE_CMD].State <> BufferStateCmd.EMPTY               ) AND
      ( Register[i].Command[ACTIVE_CMD].State <> BufferStateCmd.PROCESSED           ))
  THEN
    // copy register entry 
    TmpRegister[j] := Register[i];
    // store index of the entry from the ACR
    ExecutionOrderList[j] := i;
    // inc temporar register index
    j := j + 1; 
  END_IF
END_FOR  

// Bubble Sort to sort the priorities from the active command register
FOR i := 1 TO RegisterSize
DO
  FOR j := 1 TO RegisterSize - 1
  DO 
    // check list entry is not empty ? 
    IF (( TmpRegister[i  ].State = ActiveCommandRegisterState.IS_FREE ) OR
        ( TmpRegister[j+1].State = ActiveCommandRegisterState.IS_FREE ))
    THEN
      EXIT; 
    END_IF  

    IF (( TmpRegister[j].Command[ACTIVE_CMD].Payload[PRIORITY_IDX] AND PRIORITY_BIT_MASK ) > ( TmpRegister[j+1].Command[ACTIVE_CMD].Payload[PRIORITY_IDX] AND PRIORITY_BIT_MASK ))
    THEN    
      // swap position of register entry  
      TmpRegisterEntry := TmpRegister[j];         
      TmpRegister[j]   := TmpRegister[j+1];
      TmpRegister[j+1] := TmpRegisterEntry;
      
      // swap position of index in the Execution Order List  
      TmpIndex                := ExecutionOrderList[j];
      ExecutionOrderList[j]   := ExecutionOrderList[j+1];
      ExecutionOrderList[j+1] := TmpIndex;
    END_IF
  END_FOR 
END_FOR

// Bubble Sort to sort the Timestamp from the pre-sorted active command register
FOR i := 1 TO RegisterSize
DO
  FOR j := 1 TO RegisterSize - 1
  DO    
    // check list entry is not empty ? 
    IF (( TmpRegister[i  ].State = ActiveCommandRegisterState.IS_FREE ) OR
        ( TmpRegister[j+1].State = ActiveCommandRegisterState.IS_FREE ))
    THEN
      EXIT; 
    END_IF  

       // Priority is higher
    IF (( TmpRegister[j].Command[ACTIVE_CMD].Payload[PRIORITY_IDX] AND PRIORITY_BIT_MASK ) >= ( TmpRegister[j+1].Command[ACTIVE_CMD].Payload[PRIORITY_IDX] AND PRIORITY_BIT_MASK )) AND
       // Date is greater 
       (( TmpRegister[j].Command[ACTIVE_CMD].Timestamp.SystemDate                          >    TmpRegister[j+1].Command[ACTIVE_CMD].Timestamp.SystemDate                         ) OR 
       // Date is the same, but Time is greater
       (( TmpRegister[j].Command[ACTIVE_CMD].Timestamp.SystemDate                          =    TmpRegister[j+1].Command[ACTIVE_CMD].Timestamp.SystemDate                         ) AND 
        ( TmpRegister[j].Command[ACTIVE_CMD].Timestamp.SystemTime                          >    TmpRegister[j+1].Command[ACTIVE_CMD].Timestamp.SystemTime                         )))
    THEN    
      // swap position of register entry  
      TmpRegisterEntry := TmpRegister[j];         
      TmpRegister[j]   := TmpRegister[j+1];
      TmpRegister[j+1] := TmpRegisterEntry;
      
      // swap position of index in the Execution Order List  
      TmpIndex                := ExecutionOrderList[j];
      ExecutionOrderList[j]   := ExecutionOrderList[j+1];
      ExecutionOrderList[j+1] := TmpIndex;
    END_IF
  END_FOR 
END_FOR
END_METHOD

END_FUNCTION_BLOCK

// Library/POUs/Additional/MC_AbortMeasuringInput/MC_AbortMeasuringInputFB
/// Abort triggering of Position, measuring input
FUNCTION_BLOCK MC_AbortMeasuringInputFB EXTENDS RobotLibraryBaseExecuteFB
// ------------------------------------------------------------------------- 
//  SRCI Robot Library                                                
// ------------------------------------------------------------------------- 
//                                                                           
//  Object:      AbortMeasuringInputFB                                       
//  Author:      Thorsten Brach                                                
//  Date:        2024-06-01
//
//  Description:                                              
//   
//                                                                           
//  Copyright: 
//    (C) 2024 Thorsten Brach. All rights reserved                                                                                                                                            
//             Licensed under the MIT License.
//                                                                           
//  Disclaimer:                                                                           
//    This project is provided without any guarantee and can be used for   
//    private and commercial purposes. Any use is at the user’s 
//    own risk and responsibility.
//
// -------------------------------------------------------------------------
VAR_INPUT
  /// Command parameter 
  ParCmd          : AbortMeasuringInputParCmd;      
END_VAR
VAR_OUTPUT
  /// Command is transferred and confirmed by the RC
  CommandBuffered : BOOL;  
  /// Command output 
  OutCmd          : AbortMeasuringInputOutCmd;          
END_VAR
VAR
  /// internal copy of command parameter 
 _parCmd          : AbortMeasuringInputParCmd;
  /// command data to send
 _command         : AbortMeasuringInputSendData;
  /// response data received
 _response        : AbortMeasuringInputRecvData;      
END_VAR

SUPER^(AxesGroup := AxesGroup);

METHOD INTERNAL CheckAddParameter : BOOL
VAR_INPUT
  /// Payload pointer
  PayloadPtr : UDINT;
END_VAR
VAR
  /// Payload as byte array
  Payload    : ARRAY [1..SIZEOF(_command)] OF BYTE;
  /// Null Byte array 
  Null       : ARRAY [1..SIZEOF(_command)] OF BYTE;
  /// Data length to compare
  DataLen    : UDINT;
END_VAR
// Payload pointer must be decreased by one byte, because ADR(Payload) is already one byte !
PayloadPtr := LIMIT (0, PayloadPtr - 1, SIZEOF(Payload) -1);
// Convert command struct to payload array
SysDepMemCpy( pDest := ADR(Payload), pSrc := ADR(_command), DataLen := SIZEOF(_command));
// Calculate the data length to compare - at least one byte must be compared !
DataLen := LIMIT(1, SIZEOF(Payload) - PayloadPtr, SIZEOF(Payload)); 
// Compare Payload-Array with Null-Byte-Array
CheckAddParameter := SysDepMemCmp( pData1 := ADR(Payload) + PayloadPtr , pData2 := ADR(Null), DataLen := DataLen) <>  RobotLibraryConstants.OK ;
END_METHOD

METHOD PROTECTED CheckFunctionSupported : BOOL
VAR_IN_OUT
  /// Robot assignment of function
  AxesGroup : AxesGroup; 
END_VAR
CheckFunctionSupported := AxesGroup.State.RobotData.RCSupportedFunctions.AbortMeasuringInput;

IF ( NOT CheckFunctionSupported )
THEN
  // call base implementation for set error and create log entry
  SUPER^.CheckFunctionSupported(AxesGroup := AxesGroup);
END_IF
END_METHOD

METHOD PROTECTED CheckParameterChanged : BOOL
VAR_IN_OUT
  /// Robot assignment of function
  AxesGroup    : AxesGroup; 
END_VAR
// Check ParCmd Size is > 0, because MemCmp does not work correctly with size = 0
IF (SIZEOF(ParCmd) = 0) OR (_stepCmd = 0)
THEN 
  RETURN;
END_IF

// compare memory 
_parameterChanged := ( SysDepMemCmp(pData1 := ADR(ParCmd), pData2 := ADR(_parCmd), DataLen := SIZEOF(ParCmd)) <> RobotLibraryConstants.OK );

// check parameter valid ?
_parameterValid   := CheckParameterValid( AxesGroup := AxesGroup );

IF ((  _parameterChanged        )  AND 
    (  _parameterValid          )) OR
    (  _parameterUpdateInternal )  
THEN  
  // Create log entry for parameter changed event
  CreateLogMessagePara1 ( Timestamp   := AxesGroup.State.SystemTime,
                          MessageType := MessageType.CMD,
                          Severity    := Severity.DEBUG,
                          MessageCode := 0,
                          MessageText := 'NotifyParameterChanged Event {1}',
                          Para1       :=  '' );

  // reset internal flag for send parameter update
 _parameterUpdateInternal := FALSE;
  // update internal copy of parameters 
 _parCmd := ParCmd;
  // inc parameter sequence
 _command.ParSeq := _command.ParSeq + 1;
  // update command data  
  CommandData := CreateCommandPayload(AxesGroup := AxesGroup); // ( Access via reference to rCommandFB in ACR )
  // notify active command register 
  AxesGroup.Acyclic.ActiveCommandRegister.NotifyParameterChanged := _uniqueID;
END_IF
END_METHOD

METHOD PROTECTED CheckParameterValid : BOOL
VAR_IN_OUT
  /// Robot assignment of function
  AxesGroup : AxesGroup; 
END_VAR
CheckParameterValid := TRUE;


// Check ParCmd.MeasuringID valid ? 
IF ( ParCmd.MeasuringID < 0 )
THEN
  // Parameter not valid
  CheckParameterValid := FALSE;
  // Set error
  SetError( ErrorID := RobotLibraryErrorIdEnum.ERR_INVALID_PAR_CMD, Overwrite := TRUE ); 
  // Create log entry
  CreateLogMessagePara1 ( Timestamp   := AxesGroup.State.SystemTime,
                          MessageType := MessageType.CMD,
                          Severity    := Severity.ERROR,
                          MessageCode := ErrorID,
                          MessageText := 'Invalid Parameter ParCmd.MeasuringID = {1}',
                          Para1       := UINT_TO_STRING(ParCmd.MeasuringID));
  RETURN;                          
END_IF
END_METHOD

METHOD INTERNAL CreateCommandPayload : RobotLibraryCommandDataFB
VAR_IN_OUT
  /// Robot assignment of function
  AxesGroup : AxesGroup; 
END_VAR
VAR
  /// Parameter count
 _parameterCnt : DINT;
END_VAR
// Table 6-593: Sent CMD payload (PLC to RC) of "AbortMeasuringInput"
// --------------------------
// Header
// --------------------------
// Byte 000 : UINT  - Type HB     
// Byte 001 :       - Type LB    
// Byte 002 : USINT - Reserve | ExecutionMode
// Byte 003 : USINT - ParSeq  | Priority
// --------------------------
// Datablock
// --------------------------
// Byte 004 : UINT       - MeasuringID LW HB
// Byte 005 :            - MeasuringID LW LB
// set command parameter 
_command.CmdTyp      :=  CmdType.AbortMeasuringInput;
_command.ExecMode    :=  ExecMode;
_command.ParSeq      := _command.ParSeq;
_command.Priority    :=  Priority;
                     
_command.MeasuringID := parCmd.MeasuringID;

// copy command data to header
_cmdHeader := _command;
// call base implementation to copy header to payload buffer
CreateCommandPayload := SUPER^.CreateCommandPayload(AxesGroup := AxesGroup);


// Check parameter must be added ? 
IF ( CheckAddParameter(CreateCommandPayload.PayloadPtr))
THEN
  // add command.MeasuringID
  CreateCommandPayload.AddUint(_command.MeasuringID);
  // inc parameter counter
 _parameterCnt := _parameterCnt + 1;  
END_IF


// Create logging
CreateCommandPayloadLog(AxesGroup := AxesGroup, ParameterCnt := _parameterCnt);
END_METHOD

METHOD INTERNAL CreateCommandPayloadLog
VAR_IN_OUT
  /// Robot assignment of function
  AxesGroup : AxesGroup; 
END_VAR
VAR_INPUT
  /// Parameter count
  ParameterCnt : DINT;
END_VAR
// Create log entry for Parameter start
CreateLogMessagePara1 ( Timestamp   := AxesGroup.State.SystemTime,
                        MessageType := MessageType.CMD,
                        Severity    := Severity.DEBUG,
                        MessageCode := 0,
                        MessageText := 'Create command payload with {1} parameter(s) :',
                        Para1       := DINT_TO_STRING(ParameterCnt));
  

// Return if no parameter is remaining...
IF ( ParameterCnt = 0 ) THEN RETURN; END_IF
// dec remaining parameter(s)                        
ParameterCnt := ParameterCnt - 1;
// Create log entry for MeasuringID
CreateLogMessagePara1 ( Timestamp   := AxesGroup.State.SystemTime,
                        MessageType := MessageType.CMD,
                        Severity    := Severity.DEBUG,
                        MessageCode := 0,
                        MessageText := 'Command.MeasuringID = {1}',
                        Para1       :=  UINT_TO_STRING(_command.MeasuringID));
END_METHOD

METHOD FB_init : BOOL
VAR_INPUT
  /// if TRUE, the retain variables are initialized (warm start / cold start)
  bInitRetains : BOOL; 
  /// if TRUE, the instance afterwards gets moved into the copy code (online change)
  bInCopyCode  : BOOL;  
END_VAR
MyType := 'MC_AbortMeasuringInputFB';

ExecMode := ExecutionMode.PARALLEL;
Priority := PriorityLevel.NORMAL;
END_METHOD

METHOD PROTECTED OnExecRun : DINT
VAR_IN_OUT
  /// Robot assignment of function
  AxesGroup : AxesGroup; 
END_VAR
// call base implementation
SUPER^.OnExecRun(AxesGroup := AxesGroup);

CASE _stepCmd OF
  
  00:  IF ( _execute_R.Q ) AND ( NOT Error)
       THEN
         // Check function is supported and parameter are valid ?
         IF (( CheckFunctionSupported( AxesGroup := AxesGroup )) AND
             ( CheckParameterValid   ( AxesGroup := AxesGroup )))      
         THEN
           // set busy flag
           Busy := TRUE;
           // Reset command outputs
           SysDepMemSet(pDest := ADR(OutCmd), Value := 0, DataLen := SIZEOF(OutCmd));         
           // apply command parameter
          _parCmd := ParCmd;
           // init parameter sequence
          _command.ParSeq := 1;
           // create command data
           CommandData := CreateCommandPayload(AxesGroup := AxesGroup);
           // Add command to active command register
          _uniqueID := AxesGroup.Acyclic.ActiveCommandRegister.AddCmd( pCommandFB := ADR(THIS^ ));     
           // set timeout
           SetTimeout(PT := _timeoutCmd, rTimer := _timerCmd);
           // inc step counter
          _stepCmd := _stepCmd + 1;
         END_IF 
       END_IF


  01:  // Wait for responce received
       IF ( _responseReceived )
       THEN
         // reset response received flag
        _responseReceived := FALSE;
         // update state flags
         OnUpdateStateFlags(_response.State);
         // update state flags
         OnApplyOutCmd(_response.State);
                
         // Done, Aborted or Error ?
         IF (_response.State >= CmdMessageState.DONE )
         THEN
           // set timeout
           SetTimeout(PT := _timeoutCmd, rTimer := _timerCmd);
           // inc step counter
          _stepCmd := _stepCmd + 1; 
         END_IF
       END_IF


  02: IF ( NOT Execute)
      THEN
        Reset();
      END_IF     
ELSE
  // invalid step
  SetError( ErrorID := RobotLibraryErrorIdEnum.ERR_INVALID_STEP, Overwrite := TRUE );
END_CASE


// Reset FB
IF ( NOT Execute )
THEN
  Reset();
END_IF
END_METHOD

METHOD PROTECTED OnUpdateStateFlags
VAR_INPUT
  /// Command message state
  State : CmdMessageState;
END_VAR
// Reset State flags
Done:= FALSE;

CASE State OF

  // No operation or process is active
  CmdMessageState.EMPTY               :;
  // Created but not yet started
  CmdMessageState.CREATED             :;
  // Buffered and awaiting execution
  CmdMessageState.BUFFERED            : CommandBuffered := TRUE;
  // Buffered in planner for future execution
  CmdMessageState.BUFFERED_IN_PLANNER : CommandBuffered := TRUE;
  // Currently active and in progress
  CmdMessageState.ACTIVE              :;
  // Interrupted and awaiting continuation
  CmdMessageState.INTERRUPTED         :;
  // Requested for abort
  CmdMessageState.ABORT_REQUEST       :;
  // Successfully completed
  CmdMessageState.DONE                : Done  := TRUE;
                                        Busy  := FALSE;
  // Aborted before completion
  CmdMessageState.ABORTED             : Busy  := FALSE;
  // Encountered an error during execution
  CmdMessageState.ERROR               : Error := TRUE;
                                        Busy  := FALSE;
END_CASE
END_METHOD

METHOD INTERNAL ParseResponsePayload : DINT
VAR_INPUT
  /// Response data
  ResponseData : RobotLibraryResponseDataFB;
  /// Timestamp
  Timestamp    : SystemTime;  
END_VAR
VAR
  /// Parameter count
 _parameterCnt : DINT;
END_VAR
// Table 6-594: Received CMD payload (RC to PLC) of "AbortMeasuringInput"
// --------------------------
// Header
// --------------------------
// Byte 00 : USINT - ParSeq | State     
// Byte 01 : SINT  - AlarmMessageSeverity    
// Byte 02 : UINT  - AlarmMessageCode HB
// Byte 03 :       - AlarmMessageCode LB
// call base implementation to parse the header from payload buffer
ResponseData.PayloadPtr := SUPER^.ParseResponsePayload(ResponseData := ResponseData, Timestamp := Timestamp);

// ST-FIX F100: missing (trailing zero) bytes of the payload are 0, no values of the previous response
SysDepMemSet( pDest := ADR(_response), Value := 0, DataLen := SIZEOF(_response));

// copy parsed header to response
_response.ParSeq               := _rspHeader.ParSeq;
_response.State                := _rspHeader.State;
_response.AlarmMessageSeverity := _rspHeader.AlarmMessageSeverity;
_response.AlarmMessageCode     := _rspHeader.AlarmMessageCode;

// Create logging
ParseResponsePayloadLog(ResponseData := ResponseData, Timestamp := Timestamp, ParameterCnt := _parameterCnt);
END_METHOD

METHOD INTERNAL ParseResponsePayloadLog
VAR_INPUT
  /// Response data
  ResponseData : RobotLibraryResponseDataFB;
  /// Timestamp
  Timestamp    : SystemTime;  
  /// Parameter count
  ParameterCnt : DINT;
END_VAR
// Create log entry for Parameter start
CreateLogMessagePara1 ( Timestamp   := Timestamp,
                        MessageType := MessageType.CMD,
                        Severity    := Severity.DEBUG,
                        MessageCode := 0,
                        MessageText := '{1} parameter(s) to parse from the response data:',
                        Para1       := DINT_TO_STRING(ParameterCnt));
                        
// Return if no parameter is remaining...
IF ( ParameterCnt = 0 ) THEN RETURN; END_IF
// dec remaining parameter(s)                        
ParameterCnt := ParameterCnt - 1;
// Create log entry for no parameter 
CreateLogMessage      ( Timestamp   := Timestamp,
                        MessageType := MessageType.CMD,
                        Severity    := Severity.DEBUG,
                        MessageCode := 0,
                        MessageText := 'This command has no parameter to parse...');
END_METHOD

METHOD PROTECTED Reset : DINT
VAR_INPUT
END_VAR
Reset := SUPER^.Reset();

Done            := FALSE;
Busy            := FALSE;
CommandBuffered := FALSE;
END_METHOD

END_FUNCTION_BLOCK

// Library/POUs/Additional/MC_ActivateNextCommand/MC_ActivateNextCommandFB
/// Cancel currently active move command and continue with the next buffered command
FUNCTION_BLOCK MC_ActivateNextCommandFB EXTENDS RobotLibraryBaseExecuteFB
// ------------------------------------------------------------------------- 
//  SRCI Robot Library                                                
// ------------------------------------------------------------------------- 
//                                                                           
//  Object:      ActivateNextCommandFB                                       
//  Author:      Thorsten Brach                                                
//  Date:        2024-06-01
//
//  Description:                                              
//   
//                                                                           
//  Copyright: 
//    (C) 2024 Thorsten Brach. All rights reserved                                                                                                                                            
//             Licensed under the MIT License.
//                                                                           
//  Disclaimer:                                                                           
//    This project is provided without any guarantee and can be used for   
//    private and commercial purposes. Any use is at the user’s 
//    own risk and responsibility.
//
// -------------------------------------------------------------------------
VAR_INPUT
  /// Command parameter 
  ParCmd          : ActivateNextCommandParCmd;
  /// Processing mode
  ProcessingMode  : ProcessingMode;  
END_VAR
VAR_OUTPUT
  /// Command is transferred and confirmed by the RC
  CommandBuffered : BOOL;
  /// command results
  OutCmd          : ActivateNextCommandOutCmd;
END_VAR

VAR
  /// internal copy of command parameter 
 _parCmd          : ActivateNextCommandParCmd;
  /// command data to send
 _command         : ActivateNextCommandSendData;
  /// response data received
 _response        : ActivateNextCommandRecvData;   
  /// Trigger related EmitterID
 _emitterID       : ARRAY[0..3] OF SINT;
END_VAR

SUPER^(AxesGroup := AxesGroup);

METHOD INTERNAL CheckAddParameter : BOOL
VAR_INPUT
  /// Payload pointer
  PayloadPtr : UDINT;
END_VAR
VAR
  /// Payload as byte array
  Payload    : ARRAY [1..SIZEOF(_command)] OF BYTE;
  /// Null Byte array 
  Null       : ARRAY [1..SIZEOF(_command)] OF BYTE;
  /// Data length to compare
  DataLen    : UDINT;
END_VAR
// Payload pointer must be decreased by one byte, because ADR(Payload) is already one byte !
PayloadPtr := LIMIT (0, PayloadPtr - 1, SIZEOF(Payload) -1);
// Convert command struct to payload array
SysDepMemCpy( pDest := ADR(Payload), pSrc := ADR(_command), DataLen := SIZEOF(_command));
// Calculate the data length to compare - at least one byte must be compared !
DataLen := LIMIT(1, SIZEOF(Payload) - PayloadPtr, SIZEOF(Payload)); 
// Compare Payload-Array with Null-Byte-Array
CheckAddParameter := SysDepMemCmp( pData1 := ADR(Payload) + PayloadPtr , pData2 := ADR(Null), DataLen := DataLen) <>  RobotLibraryConstants.OK ;
END_METHOD

METHOD PROTECTED CheckFunctionSupported : BOOL
VAR_IN_OUT
  /// Robot assignment of function
  AxesGroup : AxesGroup; 
END_VAR
CheckFunctionSupported := AxesGroup.State.RobotData.RCSupportedFunctions.ActivateNextCommand;

IF ( NOT CheckFunctionSupported )
THEN
  // call base implementation for set error and create log entry
  SUPER^.CheckFunctionSupported(AxesGroup := AxesGroup);
END_IF
END_METHOD

METHOD PROTECTED CheckParameterChanged : BOOL
VAR_IN_OUT
  /// Robot assignment of function
  AxesGroup    : AxesGroup; 
END_VAR
// Check ParCmd Size is > 0, because MemCmp does not work correctly with size = 0
IF (SIZEOF(ParCmd) = 0) OR (_stepCmd = 0)
THEN 
  RETURN;
END_IF

// compare memory 
_parameterChanged := ( SysDepMemCmp(pData1 := ADR(ParCmd), pData2 := ADR(_parCmd), DataLen := SIZEOF(ParCmd)) <> RobotLibraryConstants.OK );

// check parameter valid ?
_parameterValid   := CheckParameterValid( AxesGroup := AxesGroup );

IF ((  _parameterChanged        )  AND 
    (  _parameterValid          )) OR
    (  _parameterUpdateInternal )  
THEN  
  // Create log entry for parameter changed event
  CreateLogMessagePara1 ( Timestamp   := AxesGroup.State.SystemTime,
                          MessageType := MessageType.CMD,
                          Severity    := Severity.DEBUG,
                          MessageCode := 0,
                          MessageText := 'NotifyParameterChanged Event {1}',
                          Para1       :=  '' );

  // reset internal flag for send parameter update
 _parameterUpdateInternal := FALSE;
  // update internal copy of parameters 
 _parCmd := ParCmd;
  // inc parameter sequence
 _command.ParSeq := _command.ParSeq + 1;
  // update command data  
  CommandData := CreateCommandPayload(AxesGroup := AxesGroup); // ( Access via reference to rCommandFB in ACR )
  // notify active command register 
  AxesGroup.Acyclic.ActiveCommandRegister.NotifyParameterChanged := _uniqueID;  
END_IF
END_METHOD

METHOD PROTECTED CheckParameterValid : BOOL
VAR_IN_OUT
  /// Robot assignment of function
  AxesGroup : AxesGroup; 
END_VAR

                  CheckParameterValid := TRUE;

// Check ParCmd.ProcessingMode defined ? 
// ST-FIX F122: the values between CONTINUOUS and DEACTIVATE are not defined either
IF (( ProcessingMode < ProcessingModeEnum.BUFFERED         ) OR // ST-FIX F26
    ( ProcessingMode > ProcessingModeEnum.TRIGGER_MULTIPLE ) OR
    (( ProcessingMode > ProcessingModeEnum.CONTINUOUS ) AND ( ProcessingMode < ProcessingModeEnum.DEACTIVATE )))
THEN
  // Parameter not valid
  CheckParameterValid := FALSE;
  // Set error
  SetError( ErrorID := RobotLibraryErrorIdEnum.ERR_PROCESSINGMODE_NOT_DEFINED, Overwrite := TRUE );
  // Create log entry
  CreateLogMessagePara1 ( Timestamp   := AxesGroup.State.SystemTime,
                          MessageType := MessageType.CMD,
                          Severity    := Severity.ERROR,
                          MessageCode := ErrorID,
                          MessageText := 'Invalid Parameter ParCmd.ProcessingMode = {1}',
                          Para1       := PROCESSING_MODE_TO_STRING(ProcessingMode));
  RETURN;                          
END_IF


// Check ParCmd.ProcessingMode valid ? 
IF (( ProcessingMode <> ProcessingModeEnum.PARALLEL         ) AND
    ( ProcessingMode <> ProcessingModeEnum.DEACTIVATE       ) AND
    ( ProcessingMode <> ProcessingModeEnum.TRIGGER_ONCE     ) AND
    ( ProcessingMode <> ProcessingModeEnum.TRIGGER_MULTIPLE ))
THEN
  // Parameter not valid
  CheckParameterValid := FALSE;
  // Set error
  SetError( ErrorID := RobotLibraryErrorIdEnum.ERR_PROCESSINGMODE_NOT_ALLOWED, Overwrite := TRUE );
  // Create log entry
  CreateLogMessagePara1 ( Timestamp   := AxesGroup.State.SystemTime,
                          MessageType := MessageType.CMD,
                          Severity    := Severity.ERROR,
                          MessageCode := ErrorID,
                          MessageText := 'Invalid Parameter ParCmd.ProcessingMode = {1}',
                          Para1       := PROCESSING_MODE_TO_STRING(ProcessingMode));
  RETURN;                          
END_IF


// Check ParCmd.ListenerID valid ? 
IF (( ParCmd.ListenerID <   0 ) OR 
    ( ParCmd.ListenerID > 127 ))
THEN
  // Parameter not valid
  CheckParameterValid := FALSE;
  // Set error
  SetError( ErrorID := RobotLibraryErrorIdEnum.ERR_LISTENERID_MUST_BE_POSITIVE, Overwrite := TRUE );
  // Create log entry
  CreateLogMessagePara1 ( Timestamp   := AxesGroup.State.SystemTime,
                          MessageType := MessageType.CMD,
                          Severity    := Severity.ERROR,
                          MessageCode := ErrorID,
                          MessageText := 'Invalid Parameter ParCmd.ListenerID = {1}',
                          Para1       := SINT_TO_STRING(ParCmd.ListenerID));                            
  RETURN;
END_IF

// ST-FIX F69: trigger IDs and SequenceFlag (table 7-1, 5.5.12.4, e.g. table 6-496)
IF ( CheckParameterValid ) AND ( ProcessingMode >= ProcessingModeEnum.TRIGGER_BUFFERED ) AND ( ParCmd.ListenerID = 0 )
THEN
  CheckParameterValid := FALSE;
  SetError( ErrorID := RobotLibraryErrorIdEnum.ERR_LISTENERID_MUST_BE_GREATER_THAN_ZERO, Overwrite := TRUE );
  // Create log entry
  CreateLogMessagePara1 ( Timestamp   := AxesGroup.State.SystemTime,
                          MessageType := MessageType.CMD,
                          Severity    := Severity.ERROR,
                          MessageCode := ErrorID,
                          MessageText := 'Invalid Parameter ParCmd.ListenerID = 0 with ProcessingMode = {1}',
                          Para1       := PROCESSING_MODE_TO_STRING(ProcessingMode));
  RETURN;
END_IF
IF ( CheckParameterValid ) AND ( ProcessingMode <> ProcessingModeEnum.DEACTIVATE ) AND NOT ( ProcessingMode >= ProcessingModeEnum.TRIGGER_BUFFERED ) AND ( ParCmd.ListenerID > 0 )
THEN
  CheckParameterValid := FALSE;
  SetError( ErrorID := RobotLibraryErrorIdEnum.ERR_LISTENERID_NOT_ALLOWED, Overwrite := TRUE );
  // Create log entry
  CreateLogMessagePara1 ( Timestamp   := AxesGroup.State.SystemTime,
                          MessageType := MessageType.CMD,
                          Severity    := Severity.ERROR,
                          MessageCode := ErrorID,
                          MessageText := 'Invalid Parameter ParCmd.ListenerID <> 0 with ProcessingMode = {1}',
                          Para1       := PROCESSING_MODE_TO_STRING(ProcessingMode));
  RETURN;
END_IF
END_METHOD

METHOD INTERNAL CreateCommandPayload : RobotLibraryCommandDataFB
VAR_IN_OUT
  /// Robot assignment of function
  AxesGroup : AxesGroup; 
END_VAR
VAR
  /// Parameter count
 _parameterCnt : DINT;
END_VAR
// Table 6-684: Sent CMD payload (PLC to RC) of "ActivateNextCommand"
// --------------------------
// Header
// --------------------------
// Byte 00 : UINT  - Type HB     
// Byte 01 :       - Type LB    
// Byte 02 : USINT - Reserve | ExecutionMode
// Byte 03 : USINT - ParSeq  | Priority
// --------------------------
// Datablock
// --------------------------
// Byte 04 : SINT - EmitterID[0]
// Byte 05 : SINT - EmitterID[1]
// Byte 06 : SINT - EmitterID[2]   
// Byte 07 : SINT - EmitterID[3]
// Byte 08 : SINT - ListenerID
// Byte 09 : BYTE - Reserve
// --------------------------

